(* IEC 61131-3 sources: daoli-st-library/DL_Base (part 18) *)

(* ---- FB_DL_SweepFreqGen.st ---- *)
(*
  Name        : FB_DL_SweepFreqGen
  Category    : DL_Base
  Version     : 1.0.0
  Purpose     : 频率扫描激励发生：线性/对数两模式按起止频率 + 驻留时间表逐段推进，相位逐拍积分输出瞬时频率与相位；/ Frequency sweep excitation generator: linear or logarithmic mode stepping through a dwell-time table between start and stop frequency, with per-scan phase integration
  溯源        : 借 lgf-siggen 的频率发生族待挖组织，clean-room 实现
  Boundary    : ① 起/止频率正域且相等不立（相等退化点频拒绝），越域锁存故障；
                ② 对数扫频禁对零取对数：起频下限 > 0 由正域闸保证（EXP/LN 仅作用于正比值）；
                ③ 相位积分逐拍累加防跳频突跳，相位回卷 2π 用条件减法（禁取模），回卷循环带上限守卫；
                ④ 使能撤除相位保持不归零，bRestart 上升沿显式重启回首段首相位；
                ⑤ 驻留表下标越界钳位（下标域闸）+ 非正驻留钳最小驻留常量；非有限派生频率该拍冻结保持输出；
                ⑥ 本件只出频率/相位激励量，不直接驱动脉冲输出口（属主边界，与 PulseGenerator 职责分立）。
*)
TYPE E_DL_SwpMode :
(
    eLin := 0,                               (* 线性扫频 / Linear sweep *)
    eLog := 10                               (* 对数扫频 / Logarithmic sweep *)
);
END_TYPE

TYPE E_DL_SwpState :
(
    eIdle  := 0,                             (* 未使能（相位保持） / Disabled, phase held *)
    eRun   := 10,                            (* 扫频运行 / Sweeping *)
    eFault := 90                             (* 故障锁存相 / Fault latched *)
);
END_TYPE

TYPE E_DL_SwpCause :
(
    eNone      := 0,                         (* 无故障成因 / No cause *)
    eCfgIllegal:= 1,                        (* 组态非法：频率域/步数/周期越域 / Illegal config *)
    ePhaseBad  := 2                         (* 非法相位兜底 / Illegal phase fallback *)
);
END_TYPE

FUNCTION_BLOCK FB_DL_SweepFreqGen
VAR_INPUT
    fStart  : REAL := 1.0;                   (* 起始频率，域 > 0 且不等于止频 [Hz] / Start frequency *)
    fEnd    : REAL := 100.0;                 (* 结束频率，域 > 0 且不等于起频 [Hz] / Stop frequency *)
    eMode   : E_DL_SwpMode := E_DL_SwpMode.eLin;   (* 扫频模式 / Sweep mode *)
    nSteps  : INT := 8;                      (* 驻留段数，域 2..32 [段] / Dwell step count *)
    aDwell  : ARRAY[1..32] OF TIME;          (* 各段驻留时间表（越界/非正钳位）[ms] / Dwell time table *)
    tScan   : TIME := T#10MS;                (* 扫描周期，域 > T#0S [ms] / Scan period *)
    bRepeat : BOOL := TRUE;                  (* 扫完循环重扫 [-] / Repeat sweep *)
    bEnable : BOOL := TRUE;                  (* 使能（撤除相位保持）[-] / Enable *)
    bRestart: BOOL := FALSE;                 (* 重启命令，上升沿回首段 [-] / Restart command *)
    bReset  : BOOL := FALSE;                 (* 复位命令，上升沿清故障与相位 [-] / Reset command *)
END_VAR
VAR_OUTPUT
    fFreq   : REAL;                          (* 当前瞬时频率出口 [Hz] / Instantaneous frequency outlet *)
    fPhase  : REAL;                          (* 相位累计出口（撤使能保持）[rad] / Phase accumulator outlet *)
    bSweepDone: BOOL;                        (* 单遍扫完脉冲（单拍）[-] / Sweep done pulse *)
    nSegIdx : INT;                           (* 当前段序号 [段] / Current segment index *)
    eState  : E_DL_SwpState;                 (* 状态出口 / State outlet *)
    eCause  : E_DL_SwpCause;                 (* 故障成因出口（R190 归因唯一） / Fault cause outlet *)
    bError  : BOOL;                          (* 故障锁存标志 [-] / Fault latch flag *)
END_VAR
VAR
    _eState : E_DL_SwpState := E_DL_SwpState.eIdle;  (* 内部相位（CASE 唯一写入目标） / Internal phase *)
    _eCause : E_DL_SwpCause := E_DL_SwpCause.eNone;  (* 故障成因锁存量 / Latched cause *)
    rtRestart: R_TRIG;                       (* 重启沿实例，段 0 无条件调用 / Restart edge instance *)
    rtReset : R_TRIG;                        (* 复位沿实例，段 0 无条件调用 / Reset edge instance *)
    _bFault : BOOL;                          (* 故障锁存位 / Latched fault bit *)
    _bCfgBad: BOOL;                          (* 组态非法当拍量 / Illegal config this scan *)
    _bDoneI : BOOL;                          (* 扫完脉冲内部量（统一出口映射，R187） / Done pulse internal *)
    _bFinI  : BOOL;                          (* 派生频率有限性当拍量（边界⑤） / Derived frequency finiteness *)
    _nStepsE: INT;                           (* 钳位后生效段数 [段] / Effective step count *)
    _nSegI  : INT;                           (* 内部当前段序号 [段] / Internal segment index *)
    _fDtSec : REAL;                          (* 扫描周期秒值，域 > eps [s] / Scan period seconds *)
    _fDwellS: REAL;                          (* 当前段驻留秒值（钳位后）[s] / Current dwell seconds *)
    _fTacc  : REAL;                          (* 段内驻留计时累加量 [s] / Dwell time accumulator *)
    _fFreqI : REAL;                          (* 内部瞬时频率中间量 [Hz] / Internal frequency *)
    _fPhaseI: REAL;                          (* 内部相位累计量 [rad] / Internal phase *)
    _fRatio : REAL;                          (* 对数模式频比中间量（恒正）[-] / Log mode ratio *)
    _fWrap  : INT;                           (* 相位回卷守卫计数（防死循环）[次] / Phase wrap guard *)
    _i      : INT;                           (* 驻留表下标中间量 [段] / Dwell table index *)
END_VAR
VAR CONSTANT
    DL_SWP_NMIN  : INT   := 2;               (* 段数下限（边界①域闸配套）[段] / Step count lower bound *)
    DL_SWP_NMAX  : INT   := 32;              (* 段数上限 [段] / Step count upper bound *)
    DL_SWP_EPS   : REAL  := 1.0E-6;          (* 判零容差 [-] / Epsilon *)
    DL_SWP_2PI   : REAL  := 6.2831853;       (* 相位回卷阈（2π 常量）[rad] / Phase wrap threshold *)
    DL_SWP_WRAPMAX: INT  := 64;              (* 相位回卷循环守卫上限（防死循环，边界③）[次] / Wrap loop guard *)
    DL_SWP_TDWMIN: REAL  := 0.01;            (* 最小驻留秒值（非正驻留钳位，边界⑤）[s] / Min dwell seconds *)
END_VAR

(* —— 段 0：当拍判据派生 + 实例无条件刷新（R228A） —— *)
_fDtSec := TIME_TO_LREAL(tScan) / 1000.0;                (* 扫描周期秒化（除子常量 1000） / Scan period seconds *)
_bCfgBad := (fStart <= DL_SWP_EPS) OR (fEnd <= DL_SWP_EPS)              (* 起止频率正域闸（边界①②） / Frequency positive gates *)
            OR (ABS(fStart - fEnd) < DL_SWP_EPS)                        (* 起止相等拒绝（退化点频不立，边界①） / Equal rejected *)
            OR (nSteps < DL_SWP_NMIN) OR (nSteps > DL_SWP_NMAX)         (* 段数域闸 / Step count gate *)
            OR NOT (tScan > T#0S);                                      (* 扫描周期正域闸 / Scan period gate *)
rtRestart(CLK := bRestart);                              (* 重启沿每拍必调 / Restart edge every scan *)
rtReset(CLK := bReset);                                  (* 复位沿每拍必调 / Reset edge every scan *)
_nStepsE := nSteps;                                      (* 生效段数初值 / Effective steps init *)
IF _nStepsE < DL_SWP_NMIN THEN
    _nStepsE := DL_SWP_NMIN;                             (* 段数下限钳位 / Steps lower clamp *)
END_IF
IF _nStepsE > DL_SWP_NMAX THEN
    _nStepsE := DL_SWP_NMAX;                             (* 段数上限钳位 / Steps upper clamp *)
END_IF

(* —— 段 1：单拍量预清零（R107） —— *)
_bDoneI := FALSE;                                        (* 扫完脉冲内部量预清 / Done preset *)
bSweepDone := FALSE;                                     (* 扫完脉冲出口预清 / Done outlet preset *)
_fFreqI := fFreq;                                        (* 频率中间量保持上拍（非有限拍冻结语义，边界⑤） / Frequency hold default *)

(* —— 段 2：复位沿处理（作用域：清故障 + 清相位与段序 + 迁 eIdle，R283 逐项声明） —— *)
IF rtReset.Q THEN
    _bFault := FALSE;                                    (* 清故障锁存 / Clear fault *)
    _eCause := E_DL_SwpCause.eNone;                      (* 清成因 / Clear cause *)
    _fPhaseI := 0.0;                                     (* 清相位累计 / Clear phase *)
    _nSegI := 1;                                         (* 段序回首段 / Segment to first *)
    _fTacc := 0.0;                                       (* 清驻留计时 / Clear dwell timer *)
    fFreq := 0.0;                                        (* 清频率出口 / Clear frequency outlet *)
    fPhase := 0.0;                                       (* 清相位出口 / Clear phase outlet *)
    _eState := E_DL_SwpState.eIdle;                      (* 迁未使能相 / Back to idle *)
END_IF

(* —— 段 3：组态故障锁存（锁存至复位沿，R189） —— *)
IF _bCfgBad AND NOT _bFault THEN
    _bFault := TRUE;                                     (* 锁存故障位 / Latch fault *)
    _eCause := E_DL_SwpCause.eCfgIllegal;                (* 成因：组态非法 / Cause illegal config *)
    _eState := E_DL_SwpState.eFault;                     (* 同步迁故障相 / Migrate to fault *)
END_IF

(* —— 段 4：CASE 主状态机（ELSE 兜底迁 eFault，红线 6） —— *)
CASE _eState OF
    E_DL_SwpState.eIdle:                                 (* 未使能：相位保持不归零（边界④），频率出口确定 0 / Idle *)
        fFreq := 0.0;                                    (* 失能频率出口确定值 / Disabled frequency zero *)
        IF bEnable AND NOT _bFault THEN
            _nSegI := 1;                                 (* 迁入拍段序回首段 / Segment to first *)
            _fTacc := 0.0;                               (* 驻留计时归零 / Dwell timer zero *)
            _eState := E_DL_SwpState.eRun;               (* 进入扫频相 / Enter sweeping *)
        END_IF
    E_DL_SwpState.eRun:                                  (* 扫频相：段推进 + 相位积分 / Sweeping *)
        IF NOT bEnable THEN
            _eState := E_DL_SwpState.eIdle;              (* 失能回未使能（相位保持） / Back to idle *)
        ELSE
            IF rtRestart.Q THEN
                _nSegI := 1;                             (* 显式重启回首段（边界④） / Explicit restart *)
                _fTacc := 0.0;                           (* 驻留计时归零 / Dwell timer zero *)
                _fPhaseI := 0.0;                         (* 重启相位归零 / Phase zero *)
            END_IF
            _i := _nSegI;                                (* 驻留表下标中间量 / Dwell index *)
            IF _i < 1 THEN
                _i := 1;                                 (* 下标下钳（防越界读，边界⑤） / Index lower clamp *)
            END_IF
            IF _i > DL_SWP_NMAX THEN
                _i := DL_SWP_NMAX;                       (* 下标上钳（防越界读，边界⑤） / Index upper clamp *)
            END_IF
            _fDwellS := TIME_TO_LREAL(aDwell[_i]) / 1000.0;   (* 驻留秒化（除子常量 1000） / Dwell seconds *)
            IF _fDwellS < DL_SWP_TDWMIN THEN
                _fDwellS := DL_SWP_TDWMIN;               (* 非正/过小驻留钳最小值（边界⑤） / Dwell clamp *)
            END_IF
            IF _fDtSec > DL_SWP_EPS THEN                 (* 周期秒值有效才推进（防除零/防零步进） / Period gate *)
                IF eMode = E_DL_SwpMode.eLog THEN
                    _fRatio := fEnd / fStart;            (* 对数频比（分子分母均过正域闸，边界②） / Log ratio *)
                    _fFreqI := fStart * EXP(LN(_fRatio) * INT_TO_REAL(_nSegI - 1) / INT_TO_REAL(_nStepsE - 1));   (* 几何步进频率（除子 = 段数-1 >= 1） / Geometric frequency *)
                ELSE
                    _fFreqI := fStart + (fEnd - fStart) * INT_TO_REAL(_nSegI - 1) / INT_TO_REAL(_nStepsE - 1);    (* 线性步进频率（除子 >= 1） / Linear frequency *)
                END_IF
                _bFinI := (_fFreqI = _fFreqI) AND ((_fFreqI - _fFreqI) = (_fFreqI - _fFreqI));   (* 派生频率有限性闸（边界⑤） / Derived finiteness gate *)
                IF _bFinI THEN
                    _fPhaseI := _fPhaseI + DL_SWP_2PI * _fFreqI * _fDtSec;   (* 相位逐拍积分防跳频突跳（边界③） / Phase integrate *)
                    _fWrap := 0;                         (* 回卷守卫计数清零 / Wrap guard clear *)
                    WHILE (_fPhaseI >= DL_SWP_2PI) AND (_fWrap < DL_SWP_WRAPMAX) DO   (* 条件减法回卷（禁取模，边界③） / Conditional wrap *)
                        _fPhaseI := _fPhaseI - DL_SWP_2PI;   (* 相位减 2π / Phase minus 2 pi *)
                        _fWrap := _fWrap + 1;            (* 守卫计数递进 / Guard advance *)
                    END_WHILE
                    fFreq := _fFreqI;                    (* 频率出口（有限拍派生） / Frequency outlet *)
                    fPhase := _fPhaseI;                  (* 相位出口 / Phase outlet *)
                    _fTacc := _fTacc + _fDtSec;          (* 段内驻留计时累加 / Dwell timer advance *)
                    IF _fTacc >= _fDwellS THEN           (* 驻留满迁下一段 / Dwell elapsed *)
                        _fTacc := 0.0;                   (* 驻留计时重置（R227） / Dwell timer reset *)
                        _nSegI := _nSegI + 1;            (* 段序净额 +1 / Segment advance *)
                        IF _nSegI > _nStepsE THEN        (* 末段完成 / Last segment done *)
                            _bDoneI := TRUE;             (* 扫完脉冲内部置位（R187） / Done internal *)
                            IF bRepeat THEN
                                _nSegI := 1;             (* 循环重扫回首段 / Repeat to first *)
                            ELSE
                                _nSegI := _nStepsE;      (* 单遍模式停末段（频率保持） / Hold last segment *)
                            END_IF
                        END_IF
                    END_IF
                END_IF                                   (* 非有限拍：频率/相位冻结保持上拍（边界⑤） *)
            END_IF
            nSegIdx := _nSegI;                           (* 当前段序号出口 / Segment index outlet *)
        END_IF
    E_DL_SwpState.eFault:                                (* 故障相：冻结保持末值，仅复位沿出 / Fault *)
        ;                                                (* 锁存回放（R28） / Replay from latch *)
    ELSE                                                 (* 非法相位兜底迁安全态 / Illegal phase fallback *)
        _eState := E_DL_SwpState.eFault; _bFault := TRUE;    (* 迁故障相 + 同步锁存 / To fault and latch *)
        _eCause := E_DL_SwpCause.ePhaseBad;              (* 成因：非法相位 / Cause illegal phase *)
END_CASE

(* —— 段 5：出口映射（内部 _b* → 输出单拍，R187；名实双出口，R191） —— *)
bSweepDone := _bDoneI;                                   (* 扫完脉冲单拍出口 / Done pulse outlet *)
bError := _bFault;                                       (* 故障标志镜像 / Fault flag mirror *)
eState := _eState;                                       (* 状态出口 / State outlet *)
eCause := _eCause;                                       (* 成因出口 / Cause outlet *)
END_FUNCTION_BLOCK

(* ---- FB_DL_TimerFailSafe.st ---- *)
(*
  ==================================================================
  组件名 Component  : FB_DL_TimerFailSafe
  分类   Category   : DL_Base
  复杂度 Complexity  : 轻
  版本   Version    : 1.0.0
  功能   Purpose    : 安全侧定时器。接通延时输出 bOut；当输出持续时长超过
                      tMaxHold 看门狗窗时自动回安全态 FALSE 并锁存 bTimedOut，
                      解除路径 = bIn 断电或 bReset 上升沿。安全侧赋值单点完成
                      （bOut := tonDelay.Q AND NOT _bLatch），不受本闸判定量
                      污染；与 FB_DL_ExtendedTimer 通用四模式分工互引。
  来源   Source     : T0-iec-std-wrapper（T0-2 定时器安全语义扩展）
  溯源   Origin     : IEC 61131-3 TON 标准语义的安全包装，clean-room 自研实现，
                      未复制任何厂商私有库源码。
  平台   Platform   : 纯 IEC 61131-3（Standard.library: TON / R_TRIG，无私有库）
  分工声明 Split     : 与 FB_DL_ExtendedTimer 分工——后者做通用四模式定时，
                      本件只做安全侧超时自动回退封装。
  作者   Author     : 道莅代码库 · PLC 编程专家（R59）
  ------------------------------------------------------------------
  边界 Boundary     :
                      一 安全语义：bOut 唯一赋值点为统一出口，锁存期强制 FALSE
                         （安全态），锁存解除后须 bIn 重新接通才重新计时；
                      二 组态域：tOnDelay / tMaxHold 由调用方保证为正时长，
                         本件不做二次钳制；
                      三 定时器与沿检测全部段 0 无条件周期刷新（R7）；
                      四 无全局变量、无外部变量声明、无物理地址寻址。
  修订记录 Revision  :
    2026-11-21  v1.0.0  R59 首版（批 1 · 序号 1）
  ==================================================================
*)

FUNCTION_BLOCK FB_DL_TimerFailSafe
VAR_INPUT
    bIn       : BOOL := FALSE;  // 定时条件输入，TRUE = 请求延时接通 [-] / the timing condition input, true = the on delay requested
    tOnDelay  : TIME := T#2S;   // 接通延时整定 [毫秒] / the on delay setting [millisecond]
    tMaxHold  : TIME := T#60S;  // 输出最大允许持续时长，超过自动安全态 [毫秒] / the max allowed hold duration, safe state beyond [millisecond]
    bReset    : BOOL := FALSE;  // 超时锁存复位，上升沿生效 [-] / the timeout latch reset, rising edge effective
END_VAR
VAR_OUTPUT
    bOut      : BOOL := FALSE;  // 安全侧定时输出，超时自动回 FALSE [-] / the safety side timed output, safe false on timeout
    bRun      : BOOL := FALSE;  // 延时计时进行指示 [-] / the delay timing in progress indicator
    bTimedOut : BOOL := FALSE;  // 超时锁存指示，解除 = bIn 断电或复位沿 [-] / the timeout latch indicator, released by input drop or reset edge
    bError    : BOOL := FALSE;  // 预留故障位（本件无浮点运算，恒常假）[-] / the reserved fault bit, constant false in this block
END_VAR
VAR
    _bInit   : BOOL := FALSE; // 首拍初始化标志（R310，真实使用：首拍强制安全态预置）/ the first scan flag, real use, the safe preset on first scan
    _bLatch  : BOOL := FALSE; // 超时锁存位（安全态保持源，区分于实时镜像 bTimedOut）/ the timeout latch bit, the safe state source
    rtReset  : R_TRIG;        // 复位沿检测，段 0 无条件刷新 / the reset edge, refreshed unconditionally at segment 0
    tonDelay : TON;           // 接通延时器，段 0 无条件刷新 / the on delay timer, refreshed unconditionally
    tonHold  : TON;           // 持续时长看门狗，段 0 无条件刷新 / the hold watchdog timer, refreshed unconditionally
END_VAR

// 段 0｜定时器与沿检测无条件周期刷新（禁入分支，R7）/ segment 0, the unconditional refresh
rtReset(CLK := bReset); // 复位沿 / the reset edge
tonDelay(IN := bIn AND (NOT _bLatch), PT := tOnDelay); // 接通延时，锁存期不计时 / the on delay, not timing while latched
tonHold(IN := tonDelay.Q AND (NOT _bLatch), PT := tMaxHold); // 持续看门狗，仅在输出成立期计时 / the hold watchdog, timing only while the output stands

// 段 1｜首拍初始化（R310 真实使用路径）：强制安全态预置 / segment 1, the first scan init, the safe preset
IF NOT _bInit THEN // 首拍一拍 / the first scan
    _bInit := TRUE; // 置首拍标志 / raise the first scan flag
    _bLatch := FALSE; // 锁存清零（编译缺省之上的显式安全预置）/ clear the latch explicitly
    bOut := FALSE; // 输出强制安全态 / force the output safe
END_IF

// 段 2｜超时锁存与解除（锁存解除路径 = bIn 断电沿或 bReset 上升沿，双路径可达，R188）/ segment 2, the timeout latch and release
IF tonHold.Q THEN // 看门狗窗到期：超时锁存 / the watchdog expired, latch the timeout
    _bLatch := TRUE; // 置超时锁存 / raise the timeout latch
END_IF
IF (NOT bIn) OR rtReset.Q THEN // 条件断电或复位沿 / the condition dropped or the reset edge
    _bLatch := FALSE; // 解除锁存（解除后再接通需重新计时）/ release the latch
END_IF

// 段 3｜统一出口：安全侧赋值单点完成（判定量 bIn 只经 tonDelay.Q 进入，不被闸判定量污染，边界一）/ segment 3, the unified outlet
bOut := tonDelay.Q AND (NOT _bLatch); // 输出 = 延时到 且 未超时锁存 / the output, delayed and not latched
bRun := tonDelay.IN; // 计时进行镜像 / the timing in progress mirror
bTimedOut := _bLatch; // 超时指示与锁存位同源（R191 名实双出口）/ the timeout indicator shares the latch
END_FUNCTION_BLOCK

(* ---- FB_DL_TimeWindowCheck.st ---- *)
(*==============================================================================
 * 组件名称 (Component)  : FB_DL_TimeWindowCheck
 * 所属子库 (Sublibrary) : DL_Base
 * 当前版本 (Version)    : 1.0.0
 * 兼容性   (Platform)   : CODESYS 3.5 / TwinCAT 3 / 汇川 InoProShop / Machine Expert
 *                         仅依赖 Standard.library（R_TRIG / MIN），零厂商方言
 * 分类     (Category)   : 功能块（FUNCTION_BLOCK）· 每日时间窗判定 · Level 0 DL_Base 补强件
 * 功能描述 (Function)   : 每日时间窗单一语义判定块（LGF mode 巨无霸反例的落实：
 *                         不设 MODE 参数，每周/每月/每年窗按矩阵扩产规则拆独立
 *                         块）。判定 = 本日总使能 AND 星期表当日位 AND 时刻窗。
 *                         时刻窗支持跨零点（如 22:00→06:00：t≥开 OR t<关）；
 *                         开=关视为 24h 全开（语义见段内注释）。窗口开/闭沿
 *                         单发脉冲供启停设备一次触发。当前时刻/星期由引脚注入
 *                         （零全局耦合红线：禁读 CPU 本地钟），典型与
 *                         FC_DL_DayOfWeekCalc 输出直连。
 * 开源溯源 (Origin)     : 来源标签 lgf-datetime（Siemens LGF V5.2.1 · 3.1 Date
 *                         and timer operations 章 定时开关族）。仅借鉴每日窗/
 *                         跨零点判定与星期使能表的公开行为语义；去 mode 巨无霸
 *                         化（单一语义拆块）、去 CPU 钟耦合（时间引脚注入）均
 *                         为本库独立设计决策，clean-room 重写，未复制任何源码行。
 * 本文件内含       : FUNCTION_BLOCK FB_DL_TimeWindowCheck
 * 依赖     (Depends)    : Standard.library: R_TRIG / MIN；建议上游搭配
 *                          FC_DL_DayOfWeekCalc（ISO 序星期源，引脚注入）。
 *                          不引用 DL_ 内其他实现文件。
 * 故障码表 (Error codes) : 16#0001_0202【信息级】时刻/星期参数越界（当前时刻越
 *                          界按 FALSE 处理；窗口参数越界按钳位后照常计算），
 *                          不置任何故障位（本块无故障锁存位）；0 = 无。沿用
 *                          DL_Base 既有 16#0001_xxxx 段，与 VERSION.md 故障码
 *                          表无冲突。
 * 【规格偏离留档 / R11 Deviation register】
 *   D1 规格 §4.2 引脚表未提供星期索引注入引脚，aWeekdayEnable[1..7] 表在块内
 *      无法自索引（时刻引脚不含日期信息）；按 R11 留档新增输入引脚
 *      uWeekdayNow : USINT := 1（当前星期注入，ISO 序 1=周一..7=周日，与
 *      §4.1 FC_DL_DayOfWeekCalc 输出同序同域），越界不读表并置信息级码。
 *   D2 规格引脚表 bReset 注释为「—」：本块定义其语义为上升沿清除当拍信息级码
 *      并强制重新评估窗口（日切换后防陈旧码残留），不影响窗口判定结果本身。
 * 红线自检 (Redline)    : R1 ✓ 零全局变量表与外部变量引用 ｜ R2 ✓ 零物理 IO 地址直写
 *                         R3 ✓ 纯 IEC 61131-3 ｜ R4 ✓ 越界防御+分钟折算 UINT 扩宽防溢出
 *                         R5 ✓ 全变量中英双语同行注释 ｜ R6 不适用（组合逻辑+沿检测，无状态机）
 *                         R7 ✓ 三个 R_TRIG 实例主体无条件周期刷新（严禁入分支）
 * 修订历史 (Revision)   :
 *   2026-11-15  v1.0.0  首版入库 · Round 05 · 泳道 B · 契约出处 ROUND_PLAN_R5 §4.2
 * 验收向量 (Acceptance) :
 *   V1 同日窗：On=08:00 / Off=18:00，Now=12:00 → bInWindow=TRUE；Now=07:59 /
 *      18:00 → FALSE（左闭右开）
 *   V2 跨零点窗：On=22:00 / Off=06:00，Now=23:30 或 05:59 → TRUE；Now=06:00 →
 *      FALSE；Now=21:59 → FALSE
 *   V3 24h 窗：On=Off=08:00 → 任意时刻 bInWindow=TRUE（开=关全开语义）
 *   V4 星期表：uWeekdayNow=6（周六）且 aWeekdayEnable[6]=FALSE → 不在窗，其余
 *      条件不影响；uWeekdayNow=0 或 8 → 信息级 0001_0202 且按不在窗处理
 *   V5 时刻越界：uHourNow=24 → bInWindow=FALSE + 0001_0202（当前时刻越界按
 *      FALSE 处理）；uHourOn=25 → 钳位 23 后照常计算 + 0001_0202（信息级钳位）
 *   V6 沿单发：V1 场景下 Now 由 07:59 → 08:00 当拍 bPulseOnWindowOpen=TRUE 单发；
 *      18:00 当拍 bPulseOnWindowClose=TRUE 单发
 *   V7 复位沿：越界码出现后 bReset 上升沿当拍 uErrorId 清零（触发实例无条件刷新）
 *============================================================================*)

(*==============================================================================
 * 功能块: FB_DL_TimeWindowCheck
 * 调用约定: 每个扫描周期无条件调用一次；三个 R_TRIG 实例在主体无条件周期刷新，
 *           严禁移入 IF/CASE 分支（R7）。时刻/星期由调用方每拍注入。
 *============================================================================*)
FUNCTION_BLOCK FB_DL_TimeWindowCheck
VAR_INPUT
    uHourNow        : USINT;                // 当前时刻-时（Injected local time hour）[h] 0..23，越界按不在窗处理（禁读 CPU 钟，公约 0.9）
    uMinNow         : USINT;                // 当前时刻-分（Injected local time minute）[min] 0..59
    bEnableDay      : BOOL := TRUE;         // 本日窗总使能（Day window enable），FALSE 时恒不在窗
    aWeekdayEnable  : ARRAY[1..7] OF BOOL;  // 周一~周日各日使能表（Weekday enable table），索引 1=周一（ISO 序，与 FC_DL_DayOfWeekCalc 一致）
    uWeekdayNow     : USINT := 1;           // 【偏离 D1 新增】当前星期注入（Injected weekday）1=周一..7=周日（ISO 序），越界不读表
    uHourOn         : USINT := 6;           // 窗口开启-时（Window on hour）[h] 0..23，越界钳位后照算（公约 0.2）
    uMinOn          : USINT := 0;           // 窗口开启-分（Window on minute）[min] 0..59
    uHourOff        : USINT := 22;          // 窗口关闭-时（Window off hour）[h] 0..23，支持跨零点（如 22:00→06:00）
    uMinOff         : USINT := 0;           // 窗口关闭-分（Window off minute）[min] 0..59
    bReset          : BOOL := FALSE;        // 复位（Reset）上升沿：清除当拍信息级码并重新评估（偏离 D2）
END_VAR
VAR_OUTPUT
    bInWindow           : BOOL;             // 当前处于窗口内（In window）= 本日使能 AND 星期位 AND 时刻窗
    bPulseOnWindowOpen  : BOOL;             // 窗口开启沿单发（Window open edge），TRUE 持续一拍
    bPulseOnWindowClose : BOOL;             // 窗口关闭沿单发（Window close edge），TRUE 持续一拍
    uErrorId            : UDINT;            // 信息级码（Info code）16#0001_0202 = 时刻/星期越界；0 = 无
END_VAR
VAR
    fbTrigReset     : R_TRIG;               // 复位信号上升沿检测实例（Reset edge detector）
    fbTrigOpen      : R_TRIG;               // 窗口开启沿检测实例（Window open edge detector），CLK = bInWindow
    fbTrigClose     : R_TRIG;               // 窗口关闭沿检测实例（Window close edge detector），CLK = NOT bInWindow
    uHourOnC        : USINT;                // 钳位后开启-时（Clamped on hour）[h] 0..23
    uMinOnC         : USINT;                // 钳位后开启-分（Clamped on minute）[min] 0..59
    uHourOffC       : USINT;                // 钳位后关闭-时（Clamped off hour）[h] 0..23
    uMinOffC        : USINT;                // 钳位后关闭-分（Clamped off minute）[min] 0..59
    uNowMin         : UINT;                 // 当前时刻折算分钟（Now in minutes）0..1439，USINT 域乘法越界防御
    uOnMin          : UINT;                 // 开窗时刻折算分钟（On time in minutes）0..1439
    uOffMin         : UINT;                 // 关窗时刻折算分钟（Off time in minutes）0..1439
    bTimeNowOk      : BOOL;                 // 当前时刻有效性（Now time valid）
    bWinParamOk     : BOOL;                 // 窗口参数有效性（Window params valid）
    bWeekdayOk      : BOOL;                 // 星期索引有效性（Weekday index valid）
    bTimeInWin      : BOOL;                 // 时刻窗判定结果（Time-in-window result）
    bDayOk          : BOOL;                 // 日使能合成结果（Day-enable result）
END_VAR

// -----------------------------------------------------------------------------
// 段 1｜边沿实例无条件周期刷新（R7 红线：严禁移入 IF/CASE 分支）
// -----------------------------------------------------------------------------
fbTrigReset(CLK := bReset);                 // 复位沿检测

// -----------------------------------------------------------------------------
// 段 2｜有效性判定与信息级码准备（信息级 0001_0202 只进 uErrorId，本块无故障位）
// -----------------------------------------------------------------------------
uErrorId := 16#0000_0000;                   // 每拍重算信息级码
bTimeNowOk  := (uHourNow <= 23) AND (uMinNow <= 59);               // 当前时刻域检查
bWinParamOk := (uHourOn <= 23) AND (uMinOn <= 59)
            AND (uHourOff <= 23) AND (uMinOff <= 59);          // 窗口参数域检查
bWeekdayOk  := (uWeekdayNow >= 1) AND (uWeekdayNow <= 7);      // 星期索引域检查（ISO 1..7）
IF NOT bTimeNowOk THEN
    uErrorId := 16#0001_0202;               // 当前时刻越界：按不在窗处理（引脚注释基线）
END_IF
IF NOT bWinParamOk THEN
    uErrorId := 16#0001_0202;               // 窗口参数越界：钳位后照常计算（公约 0.2）
END_IF
IF NOT bWeekdayOk THEN
    uErrorId := 16#0001_0202;               // 星期索引越界：不读表，按不在窗处理
END_IF

// -----------------------------------------------------------------------------
// 段 3｜窗口参数钳位（信息级钳位，钳位后继续计算，不中断扫描）
// -----------------------------------------------------------------------------
uHourOnC  := MIN(uHourOn, 23);              // 开启-时钳位 [h]
uMinOnC   := MIN(uMinOn, 59);               // 开启-分钳位 [min]
uHourOffC := MIN(uHourOff, 23);             // 关闭-时钳位 [h]
uMinOffC  := MIN(uMinOff, 59);              // 关闭-分钳位 [min]

// -----------------------------------------------------------------------------
// 段 4｜分钟折算（USINT×60 最大 1380 超 USINT 域，先扩宽 UINT 再运算防越界）
// -----------------------------------------------------------------------------
uOnMin := uHourOnC;                         // USINT → UINT 隐式扩宽
uOnMin := (uOnMin * 60) + uMinOnC;          // 开窗分钟 [min] 0..1439
uOffMin := uHourOffC;                       // USINT → UINT 隐式扩宽
uOffMin := (uOffMin * 60) + uMinOffC;       // 关窗分钟 [min] 0..1439
IF bTimeNowOk THEN
    uNowMin := uHourNow;                    // USINT → UINT 隐式扩宽
    uNowMin := (uNowMin * 60) + uMinNow;    // 当前分钟 [min] 0..1439
ELSE
    uNowMin := 0;                           // 时刻越界：折算值弃用，结果由 bTimeNowOk 门控
END_IF

// -----------------------------------------------------------------------------
// 段 5｜时刻窗判定（跨零点支持；开=关视为 24h 全开——语义：本日整日放行）
// -----------------------------------------------------------------------------
IF uOnMin > uOffMin THEN
    bTimeInWin := (uNowMin >= uOnMin) OR (uNowMin < uOffMin);   // 跨零点窗：t≥开 OR t<关（如 22:00→06:00）
ELSIF uOnMin < uOffMin THEN
    bTimeInWin := (uNowMin >= uOnMin) AND (uNowMin < uOffMin);  // 同日窗：开≤t<关（左闭右开）
ELSE
    bTimeInWin := TRUE;                                          // 开=关：24h 全开（每日窗单一语义特例）
END_IF

// -----------------------------------------------------------------------------
// 段 6｜日使能合成（星期越界不读表，防数组越界，R4）
// -----------------------------------------------------------------------------
IF bWeekdayOk THEN
    bDayOk := bEnableDay AND aWeekdayEnable[uWeekdayNow];       // 总使能 AND 当日星期位（索引 1..7 已校验）
ELSE
    bDayOk := FALSE;                        // 星期索引越界：按不在窗处理
END_IF

// -----------------------------------------------------------------------------
// 段 7｜总判定：当前时刻越界按 FALSE 处理；窗口参数已钳位故不再门控结果
// -----------------------------------------------------------------------------
bInWindow := bDayOk AND bTimeNowOk AND bTimeInWin;              // 在窗 = 日使能 AND 时刻有效 AND 时刻窗

// -----------------------------------------------------------------------------
// 段 8｜窗口开/闭沿单发（实例无条件周期刷新，沿输出各持续一拍）
// -----------------------------------------------------------------------------
fbTrigOpen(CLK := bInWindow);               // 开启沿检测
fbTrigClose(CLK := NOT bInWindow);          // 关闭沿检测（取反 CLK）
bPulseOnWindowOpen  := fbTrigOpen.Q;        // 开启沿单发输出
bPulseOnWindowClose := fbTrigClose.Q;       // 关闭沿单发输出

// -----------------------------------------------------------------------------
// 段 9｜复位沿消费：清除当拍信息级码（触发实例已在段 1 无条件刷新，偏离 D2）
// -----------------------------------------------------------------------------
IF fbTrigReset.Q THEN
    uErrorId := 16#0000_0000;               // 复位沿当拍清信息级码（下一拍重新评估）
END_IF

END_FUNCTION_BLOCK

(* ---- FB_DL_TofEx.st ---- *)
(*==============================================================================
 * 组件名称 (Component)  : FB_DL_TofEx
 * 所属子库 (Sublibrary) : DL_Base
 * 当前版本 (Version)    : 1.0.0
 * 兼容性   (Platform)   : CODESYS 3.5 / TwinCAT 3 / 汇川 InoProShop / Machine Expert
 *                         仅依赖 Standard.library（TOF），零厂商方言
 * 功能描述 (Function)   : 断开延时定时器防御包装。内部委托 IEC 61131-3 标准 TOF
 *                         实例完成计时内核，外围提供 PT 负值钳位、首扫语义统一
 *                         （首扫 bIN=FALSE 时 bQ 必为 FALSE）与跨段语义直通。
 * 溯源     (Origin)     : IEC 61131-3 标准语义的道莅防御性实现
 *                         （接口语义由 IEC 61131-3 定义，clean-room 重写，
 *                         参考公开标准条款）
 * 码位     (Diag Codes) : 信息级占用区间 16#0001_0150（本件独占，仅此一码）
 *                         16#0001_0150 = tPT 为负值，已钳位为 T#0s（信息级，
 *                         钳位属正常防御行为，不置故障）
 * 类型裁定 (Type Note)  : 码位段 16#0001_xxxx 为全库共享 32 位段，WORD 容量不足，
 *                         故 uDiag 采用 UDINT 承载（与库内 uErrorId : UDINT 惯例一致）
 * 依赖     (Depends)    : 无 DL_ 内部依赖；Standard.library: TOF
 * 红线自检 (Redline)    : R1 ✓ 零全局变量与外部变量引用 ｜ R2 ✓ 零物理 IO 地址直写
 *                         R3 ✓ 纯 IEC 61131-3 ｜ R4 ✓ PT 钳位+除零/越界无涉
 *                         R5 ✓ 全变量中英双语同行注释 ｜ R6 N/A（无顺序状态机，见下）
 *                         R7 ✓ TOF 实例主体无条件周期刷新
 * 说明     (Note)       : R6 标注 N/A —— 本组件为单步延时逻辑，不存在顺序状态机，
 *                         无 CASE 可写；唯一状态即"延时中/直通"，以本节说明
 *                         替代 ELSE 兜底，符合"无状态机则标注 N/A"口径。
 * 防御行为声明 (Defense): ① tPT < T#0s 时钳位为 T#0s 并置信息码 16#0001_0150
 *                           （部分平台负 TIME 行为未定义，本库统一钳 0）；
 *                         ② 首扫语义统一：首扫 bIN=FALSE 时 bQ 必为 FALSE、tET=T#0s
 *                           ——由内建 TOF 标准行为（Q 随 IN 直通 + 断开延时）保证，
 *                           部分平台首扫假触发差异在包装层被标准实例天然屏蔽；
 *                         ③ bIN 接通当拍 tET 归零、bQ 立即 TRUE（IEC TOF 标准语义，
 *                           包装层不重实现）。
 * 修订历史 (Revision)   :
 *   2026-11-16  v1.0.0  首版入库（R14 批 2 · T0 快车道）
 *============================================================================*)
FUNCTION_BLOCK FB_DL_TofEx
VAR_INPUT
    bIN : BOOL;   // 定时输入，TRUE 直通输出，FALSE 起断开延时 / Timing input, TRUE passes through, FALSE starts the off-delay
    tPT : TIME;   // 预置延时 [ms]，负值将被钳位为 T#0s / Preset delay [ms], negative values are clamped to T#0s
END_VAR
VAR_OUTPUT
    bQ    : BOOL;   // 输出，bIN 断开并持续 tPT 后变 FALSE / Output, goes FALSE after bIN held FALSE for tPT
    tET   : TIME;   // 已计时 [ms]，bIN 接通当拍归零 / Elapsed time [ms], zeroed on the scan bIN rises
    uDiag : UDINT;  // 诊断字，16#0001_0150=tPT 负值已钳 0，0=无诊断事件 / Diag word, 16#0001_0150=negative tPT clamped to 0, 0=no diag event
END_VAR
VAR
    fbTof    : TOF;   // 内建断开延时实例，承担计时内核 / Built-in TOF instance, owns the timing kernel
    tPTClamp : TIME;  // 钳位后的预置延时 [ms]，喂给内建实例 / Clamped preset delay [ms], fed to the built-in instance
    xInit    : BOOL;  // 首扫初始化标志，FALSE=尚未完成上电初始化 / First-scan init flag, FALSE = power-on init not yet done
END_VAR

(*------------------------------------------------------------------------------
 * 段 1｜首扫初始化（历史教训④口径）：置于逻辑最前，首扫不产假 bQ
 *      First-scan init (lesson 4): placed at the very front, no false bQ on first scan
 *-----------------------------------------------------------------------------*)
IF NOT xInit THEN
    xInit    := TRUE;    // 置初始化完成标志 / Mark init as done
    tPTClamp := T#0s;    // 首扫钳位值归零，避免未初始化喂入 / Zero the clamp value on first scan, no uninitialized feed
    uDiag    := 16#0000_0000;  // 首扫诊断字清零 / Clear diag word on first scan
END_IF

(*------------------------------------------------------------------------------
 * 段 2｜PT 域校验与钳位：负 TIME 在部分平台行为未定义，统一钳 0 并置信息码；
 *      写入点排序审计（历史教训⑦）：本件诊断字仅有"置码/清码"单一分支对，
 *      无复位类与置位类竞态，排序安全
 *      PT domain check and clamp: negative TIME is undefined on some platforms,
 *      unified clamp to 0 with an informational code
 *-----------------------------------------------------------------------------*)
IF tPT < T#0s THEN
    tPTClamp := T#0s;        // 负值钳位为 0 [ms] / Clamp negative to 0 [ms]
    uDiag    := 16#0001_0150;  // 信息码：PT 负值已钳 0 / Informational: negative PT clamped to 0
ELSE
    tPTClamp := tPT;         // 域内直通 / In-domain pass-through
    uDiag    := 16#0000_0000;  // 无诊断事件，清码 / No diag event, clear code
END_IF

(*------------------------------------------------------------------------------
 * 段 3｜无条件刷新区（红线 R7）：TOF 实例严禁进入任何 IF / CASE 分支；
 *      首扫 bIN=FALSE → bQ=FALSE 与"接通当拍 ET 归零"均由内建标准语义保证
 *      Unconditional refresh zone (red line R7): no instance call inside IF / CASE;
 *      first-scan bQ=FALSE with bIN=FALSE and ET zeroing on bIN rise are both
 *      guaranteed by the built-in TOF standard behavior
 *-----------------------------------------------------------------------------*)
fbTof(IN := bIN, PT := tPTClamp);  // 每扫描周期无条件喂入输入与钳位后 PT / Feed input and clamped PT unconditionally every scan

(*------------------------------------------------------------------------------
 * 段 4｜输出直通：bQ/tET 逐拍镜像内建实例输出，包装层不重实现计时内核
 *      Output pass-through: bQ/tET mirror the built-in outputs scan by scan;
 *      the wrapper never re-implements the timing kernel
 *-----------------------------------------------------------------------------*)
bQ  := fbTof.Q;   // 输出直通 / Output pass-through
tET := fbTof.ET;  // 已计时 [ms] 直通 / Elapsed time [ms] pass-through
END_FUNCTION_BLOCK

(* ---- FB_DL_ToggleButtonBank.st ---- *)
(*
  FB_DL_ToggleButtonBank  —  多路启停按钮组解算 / Multi-channel toggle button bank solver
  分类 Category : DL_Base
  码位 Code     : 16#01_0_01
  版本 Version  : 1.0.0
  来源 Source   : t1-5-tcopen — IEC 61131-3 标准语义的道莅防御性实现
  溯源 Origin   : TCopen 按钮组/选择器公开语义借鉴，clean-room 实现，未复制任何源码行
  功能 Function : 1) 三种解算模式：Toggle 单按钮逐通道翻转锁存 / SingleAct 双按钮点动直通 / Selector3 三位置选择互斥；
                  2) Selector3 通道互斥：新通道置位时旧通道清零；同拍多键按「低通道号优先」并置信息码（不静默双通）；
                  3) 失电来电恢复策略 eRestorePolicy：Hold 保持（RETAIN 语义由上层承载）/ Reset 全清 / Pulse 上电首拍单周期 TRUE；
                  4) nActiveChannel 输出当前活动通道（0 = 无，1..n = 最低活动通道号，Selector3 即唯一互斥通道）。
  边界 Boundary : ① uChannelCount = 0 或 > nMaxCh 判组态错 bCfgFault，全输出 FALSE（安全侧）；
                  ② 8 路 R_TRIG 在主周期无条件刷新（调用语句不置于 IF/CASE 内，R182）；
                  ③ SingleAct 点动直通不锁存：输出 = 按钮实时电平（松开即断，无保持）；
                  ④ 解除式自证：bCfgFault 解除 = 下一拍 uChannelCount 落回合法域（每拍重算，无锁存）；
                  ⑤ Pulse 脉冲语义：仅上电首拍 abOut 全 TRUE 一个 PLC 周期，第二拍起恢复正常解算（注释标明，防误用为持续使能）。
  依赖 Depends  : 仅 Standard.library（R_TRIG）；枚举 E_DL_BtnMode / E_DL_RestorePolicy 随本件发布
  码表 Error codes（本件格 01_0_01，子码步进 +0x100）:
    16#0001_0101 信息级：Selector3 同拍多键，低通道号优先（不置故障）
    16#0001_0201 故障级：组态非法 uChannelCount = 0 或超数组上界
    16#0001_0301 信息级：Pulse 恢复策略上电首拍单周期脉冲（不置故障）

  修订历史 Revision :
    2026-11-18  v1.0.0  R38 首版
*)

TYPE E_DL_BtnMode :
(
    eToggle    := 0,   // 单按钮翻转锁存 / Single-button toggle with latch
    eSingleAct := 1,   // 点动直通（不锁存）/ Momentary passthrough, no latch
    eSelector3 := 2    // 三位置选择互斥 / Three-position selector, mutually exclusive
);
END_TYPE

TYPE E_DL_RestorePolicy :
(
    eHold  := 0,   // 上电保持断电前状态（RETAIN 由上层承载）/ Hold pre-power-loss state, retainment owned upstream
    eReset := 1,   // 上电全清零 / Clear all outputs at power-up
    ePulse := 2    // 上电首拍单周期 TRUE / Single-scan TRUE pulse at power-up
);
END_TYPE

FUNCTION_BLOCK FB_DL_ToggleButtonBank
VAR_INPUT
    abBtn          : ARRAY[0..7] OF BOOL;   // 按钮输入组 [0..nMaxCh-1] / Button inputs
    uChannelCount  : INT;                   // 有效通道数 [路]，域 1..nMaxCh / Valid channel count
    eMode          : E_DL_BtnMode;          // 解算模式 / Solver mode
    eRestorePolicy : E_DL_RestorePolicy;    // 失电来电恢复策略 / Power-restore policy
END_VAR
VAR_OUTPUT
    abOut          : ARRAY[0..7] OF BOOL;   // 通道输出组 / Channel outputs
    nActiveChannel : INT;                   // 活动通道号（0 = 无，1..n 最低活动）/ Active channel, 0 = none
    bCfgFault      : BOOL;                  // 组态非法（每拍重算）/ Configuration fault, recomputed
    nErrId         : UDINT;                 // 事件码，0 = 无事件 / Event code, 0 = none
END_VAR
VAR
    artBtn     : ARRAY[0..7] OF R_TRIG;     // 逐通道按钮上升沿，段 0 无条件刷新 / Per-channel rising edges
    _abState   : ARRAY[0..7] OF BOOL;       // Toggle 模式锁存状态 / Toggle latched states
    _bFirstScan: BOOL := TRUE;              // 上电首拍标志 / First-scan-after-power-up flag
    _bSimulKey : BOOL;                      // 同拍多键标志（本拍重算）/ Simultaneous keys flag
    _k         : INT;                       // 循环计数器 / Loop counter
END_VAR
VAR CONSTANT
    nMaxCh : INT := 8;                      // 数组上界 [路] / Array upper bound
END_VAR

(* —— 段 0：R_TRIG 无条件周期刷新（R182：调用语句不得置于 IF/CASE 内） —— *)
FOR _k := 0 TO (nMaxCh - 1) DO
    artBtn[_k](CLK := abBtn[_k]);           // 逐通道上升沿，每拍必调
END_FOR

(* —— 段 1：单拍量预清零 —— *)
nErrId     := 16#0000_0000;               // 事件码缺省无事件
_bSimulKey := FALSE;                      // 多键标志预清零
FOR _k := 0 TO (nMaxCh - 1) DO
    abOut[_k] := FALSE;                   // 输出缺省 FALSE（安全侧缺省，段 4 单点置位）
END_FOR
nActiveChannel := 0;                      // 活动通道缺省无

(* —— 段 2：组态域闸（uChannelCount 全覆盖，每拍重算） —— *)
IF (uChannelCount <= 0) OR (uChannelCount > nMaxCh) THEN
    bCfgFault := TRUE;                    // 组态非法：全输出维持 FALSE（段 1 已清）
    nErrId    := 16#0001_0201;            // 故障级：组态非法
ELSE
    bCfgFault := FALSE;                   // 解除式自证：下一拍通道数合法即解除
END_IF

(* —— 段 3：上电首拍恢复策略（仅在组态合法时生效） —— *)
IF (NOT bCfgFault) AND _bFirstScan THEN
    CASE eRestorePolicy OF

    E_DL_RestorePolicy.eHold:
        ;                                  // 保持：_abState 维持 RETAIN 语义值（上层持久化承载）
    E_DL_RestorePolicy.eReset:
        FOR _k := 0 TO (nMaxCh - 1) DO
            _abState[_k] := FALSE;         // 上电全清
        END_FOR
    E_DL_RestorePolicy.ePulse:
        FOR _k := 0 TO (nMaxCh - 1) DO
            abOut[_k] := TRUE;             // 脉冲语义：置位 1 个 PLC 周期（规格强制，防误用为持续使能）
        END_FOR
        nErrId := 16#0001_0301;            // 信息级：Pulse 上电单拍脉冲
    ELSE
        nErrId := 16#0001_0201;            // 未知恢复策略按组态错兜底（安全侧全 FALSE）
        bCfgFault := TRUE;
    END_CASE
END_IF
_bFirstScan := FALSE;                     // 首拍标志自清

(* —— 段 4：三模式解算（组态合法才执行） —— *)
IF NOT bCfgFault THEN
    CASE eMode OF

    E_DL_BtnMode.eToggle:
        FOR _k := 0 TO (uChannelCount - 1) DO
            IF artBtn[_k].Q THEN
                _abState[_k] := NOT _abState[_k];   // 单按钮翻转锁存
            END_IF
            abOut[_k] := _abState[_k];              // 输出锁存态
        END_FOR

    E_DL_BtnMode.eSingleAct:
        FOR _k := 0 TO (uChannelCount - 1) DO
            abOut[_k] := abBtn[_k];                 // 点动直通：输出 = 按钮实时电平，松开即断
        END_FOR

    E_DL_BtnMode.eSelector3:
        FOR _k := 0 TO (uChannelCount - 1) DO
            IF abBtn[_k] THEN
                IF nActiveChannel = 0 THEN
                    nActiveChannel := _k + 1;       // 记录最低按下的通道号（低通道号优先）
                ELSE
                    _bSimulKey := TRUE;             // 同拍多键：置信息码（不做静默双通）
                END_IF
            END_IF
        END_FOR
        IF _bSimulKey THEN
            nErrId := 16#0001_0101;                 // 信息级：同拍多键，低通道号优先
        END_IF
        IF nActiveChannel > 0 THEN
            FOR _k := 0 TO (uChannelCount - 1) DO
                _abState[_k] := (_k = (nActiveChannel - 1));   // 互斥：仅选中通道保持
                abOut[_k] := _abState[_k];
            END_FOR
        ELSE
            FOR _k := 0 TO (uChannelCount - 1) DO
                _abState[_k] := FALSE;              // 无键按下：互斥组全清
            END_FOR
        END_IF

    ELSE
        bCfgFault := TRUE;                          // 未知模式兜底：全 FALSE 安全侧
        nErrId := 16#0001_0201;                     // 故障级：组态非法（模式越界并入组态错）
    END_CASE
END_IF

(* —— 段 5：活动通道出口（Toggle/SingleAct 取最低活动通道） —— *)
IF (eMode = E_DL_BtnMode.eToggle) OR (eMode = E_DL_BtnMode.eSingleAct) THEN
    nActiveChannel := 0;                            // 缺省无
    FOR _k := 0 TO (uChannelCount - 1) DO
        IF abOut[_k] THEN
            nActiveChannel := _k + 1;               // 最低活动通道号
            EXIT;                                    // 找到即止
        END_IF
    END_FOR
END_IF

END_FUNCTION_BLOCK

(* ---- FB_DL_TonEx.st ---- *)
(*==============================================================================
 * 组件名称 (Component)  : FB_DL_TonEx
 * 所属子库 (Sublibrary) : DL_Base
 * 当前版本 (Version)    : 1.0.0
 * 兼容性   (Platform)   : CODESYS 3.5 / TwinCAT 3 / 汇川 InoProShop / Machine Expert
 *                         仅依赖 Standard.library（TON），零厂商方言
 * 功能描述 (Function)   : 接通延时定时器防御包装。内部委托 IEC 61131-3 标准 TON
 *                         实例完成计时内核，外围提供 PT 负值钳位与跨段输入断开
 *                         语义统一（bIN 断开当拍 ET 归零、bQ 立即 FALSE）。
 * 溯源     (Origin)     : IEC 61131-3 标准语义的道莅防御性实现
 *                         （接口语义由 IEC 61131-3 定义，clean-room 重写，
 *                         参考公开标准条款）
 * 码位     (Diag Codes) : 信息级占用区间 16#0001_014F（本件独占，仅此一码）
 *                         16#0001_014F = tPT 为负值，已钳位为 T#0s（信息级，
 *                         钳位属正常防御行为，不置故障）
 * 类型裁定 (Type Note)  : 码位段 16#0001_xxxx 为全库共享 32 位段，WORD 容量不足，
 *                         故 uDiag 采用 UDINT 承载（与库内 uErrorId : UDINT 惯例一致）
 * 依赖     (Depends)    : 无 DL_ 内部依赖；Standard.library: TON
 * 红线自检 (Redline)    : R1 ✓ 零全局变量与外部变量引用 ｜ R2 ✓ 零物理 IO 地址直写
 *                         R3 ✓ 纯 IEC 61131-3 ｜ R4 ✓ PT 钳位+除零/越界无涉
 *                         R5 ✓ 全变量中英双语同行注释 ｜ R6 N/A（无顺序状态机，见下）
 *                         R7 ✓ TON 实例主体无条件周期刷新
 * 说明     (Note)       : R6 标注 N/A —— 本组件为单步延时逻辑，不存在顺序状态机，
 *                         无 CASE 可写；非法状态不可能出现（唯一状态即"计时/直通"），
 *                         故以本节说明替代 ELSE 兜底，符合"无状态机则标注 N/A"口径。
 * 防御行为声明 (Defense): ① tPT < T#0s 时钳位为 T#0s 并置信息码 16#0001_014F
 *                           （部分平台负 TIME 行为未定义，本库统一钳 0）；
 *                         ② 跨段输入断开语义统一：bIN 断开当拍 tET 归零、bQ 立即
 *                           FALSE（由内建 TON 标准语义保证，包装层不重实现）；
 *                         ③ 首扫 bIN=TRUE 允许正常计时（TON 标准语义）但不产假 bQ
 *                           （首拍 ET 从 0 起步，bQ 天然 FALSE，无需额外抑制）。
 * 修订历史 (Revision)   :
 *   2026-11-16  v1.0.0  首版入库（R14 批 1 · T0 快车道）
 *============================================================================*)
FUNCTION_BLOCK FB_DL_TonEx
VAR_INPUT
    bIN : BOOL;   // 定时输入，TRUE 起计时，FALSE 立即复位计时 / Timing input, TRUE starts timing, FALSE resets immediately
    tPT : TIME;   // 预置延时 [ms]，负值将被钳位为 T#0s / Preset delay [ms], negative values are clamped to T#0s
END_VAR
VAR_OUTPUT
    bQ    : BOOL;   // 延时到输出，bIN 保持 TRUE 达 tPT 后置位 / Delay-elapsed output, set after bIN held TRUE for tPT
    tET   : TIME;   // 已计时 [ms]，bIN 断开当拍归零 / Elapsed time [ms], zeroed on the scan bIN drops
    uDiag : UDINT;  // 诊断字，16#0001_014F=tPT 负值已钳 0，0=无诊断事件 / Diag word, 16#0001_014F=negative tPT clamped to 0, 0=no diag event
END_VAR
VAR
    fbTon    : TON;   // 内建接通延时实例，承担计时内核 / Built-in TON instance, owns the timing kernel
    tPTClamp : TIME;  // 钳位后的预置延时 [ms]，喂给内建实例 / Clamped preset delay [ms], fed to the built-in instance
    xInit    : BOOL;  // 首扫初始化标志，FALSE=尚未完成上电初始化 / First-scan init flag, FALSE = power-on init not yet done
END_VAR

(*------------------------------------------------------------------------------
 * 段 1｜首扫初始化（历史教训⑤口径）：置于逻辑最前，禁止"初值置位后同步清零"反模式
 *      First-scan init (lesson 5): placed at the very front of the logic body
 *-----------------------------------------------------------------------------*)
IF NOT xInit THEN
    xInit    := TRUE;    // 置初始化完成标志 / Mark init as done
    tPTClamp := T#0s;    // 首扫钳位值归零，避免未初始化喂入 / Zero the clamp value on first scan, no uninitialized feed
    uDiag    := 16#0000_0000;  // 首扫诊断字清零 / Clear diag word on first scan
END_IF

(*------------------------------------------------------------------------------
 * 段 2｜PT 域校验与钳位：负 TIME 在部分平台行为未定义，统一钳 0 并置信息码；
 *      写入点排序（历史教训⑩）：本件诊断字仅有"置码 / 清码"单一分支对，无
 *      复位类与置位类竞态，排序安全
 *      PT domain check and clamp: negative TIME is undefined on some platforms,
 *      unified clamp to 0 with an informational code
 *-----------------------------------------------------------------------------*)
IF tPT < T#0s THEN
    tPTClamp := T#0s;        // 负值钳位为 0 [ms] / Clamp negative to 0 [ms]
    uDiag    := 16#0001_014F;  // 信息码：PT 负值已钳 0 / Informational: negative PT clamped to 0
ELSE
    tPTClamp := tPT;         // 域内直通 / In-domain pass-through
    uDiag    := 16#0000_0000;  // 无诊断事件，清码 / No diag event, clear code
END_IF

(*------------------------------------------------------------------------------
 * 段 3｜无条件刷新区（红线 R7）：TON 实例严禁进入任何 IF / CASE 分支；
 *      bIN 断开当拍 ET 归零、bQ 立即 FALSE 的跨段统一语义由内建 TON 标准行为保证
 *      Unconditional refresh zone (red line R7): no instance call inside IF / CASE;
 *      the unified drop-out semantics (ET zeroed and bQ FALSE on the scan bIN
 *      drops) is guaranteed by the built-in TON standard behavior
 *-----------------------------------------------------------------------------*)
fbTon(IN := bIN, PT := tPTClamp);  // 每扫描周期无条件喂入输入与钳位后 PT / Feed input and clamped PT unconditionally every scan

(*------------------------------------------------------------------------------
 * 段 4｜输出直通：bQ/tET 逐拍镜像内建实例输出，包装层不重实现计时内核
 *      Output pass-through: bQ/tET mirror the built-in outputs scan by scan;
 *      the wrapper never re-implements the timing kernel
 *-----------------------------------------------------------------------------*)
bQ  := fbTon.Q;   // 延时到输出直通 / Delay-elapsed output pass-through
tET := fbTon.ET;  // 已计时 [ms] 直通 / Elapsed time [ms] pass-through
END_FUNCTION_BLOCK

(* ---- FB_DL_TpEx.st ---- *)
(*==============================================================================
 * 组件名称 (Component)  : FB_DL_TpEx
 * 所属子库 (Sublibrary) : DL_Base
 * 当前版本 (Version)    : 1.0.0
 * 兼容性   (Platform)   : CODESYS 3.5 / TwinCAT 3 / 汇川 InoProShop / Machine Expert
 *                         仅依赖 Standard.library（TP），零厂商方言
 * 功能描述 (Function)   : 脉冲定时器防御包装。内部委托 IEC 61131-3 标准 TP 实例
 *                         完成计时内核，外围提供 PT 负值钳位，并把"不可重触发"
 *                         语义在头注释显式写死。
 * 溯源     (Origin)     : IEC 61131-3 标准语义的道莅防御性实现
 *                         （接口语义由 IEC 61131-3 定义，clean-room 重写，
 *                         参考公开标准条款）
 * 码位     (Diag Codes) : 信息级占用区间 16#0001_0151（本件独占，仅此一码）
 *                         16#0001_0151 = tPT 为负值，已钳位为 T#0s（信息级，
 *                         钳位属正常防御行为，不置故障）
 * 类型裁定 (Type Note)  : 码位段 16#0001_xxxx 为全库共享 32 位段，WORD 容量不足，
 *                         故 uDiag 采用 UDINT 承载（与库内 uErrorId : UDINT 惯例一致）
 * 依赖     (Depends)    : 无 DL_ 内部依赖；Standard.library: TP
 * 红线自检 (Redline)    : R1 ✓ 零全局变量与外部变量引用 ｜ R2 ✓ 零物理 IO 地址直写
 *                         R3 ✓ 纯 IEC 61131-3 ｜ R4 ✓ PT 钳位+除零/越界无涉
 *                         R5 ✓ 全变量中英双语同行注释 ｜ R6 N/A（无顺序状态机，见下）
 *                         R7 ✓ TP 实例主体无条件周期刷新
 * 说明     (Note)       : R6 标注 N/A —— 本组件为单步脉冲逻辑，不存在顺序状态机，
 *                         无 CASE 可写；唯一状态即"脉冲中/待触发"，以本节说明
 *                         替代 ELSE 兜底，符合"无状态机则标注 N/A"口径。
 * 防御行为声明 (Defense): ① tPT < T#0s 时钳位为 T#0s 并置信息码 16#0001_0151
 *                           （部分平台负 TIME 行为未定义，本库统一钳 0，
 *                           PT=0 时脉冲退化为单扫描周期宽度）；
 *                         ② 不可重触发语义显式化（IEC TP 标准语义，多平台实现
 *                           有偏差，此处以标准实例写死）：计时进行中 bIN 再次
 *                           触发不延长、不重启当前脉冲，必须等当前脉冲结束；
 *                         ③ R24 教训落实：本件不存在任何"实例调用前的自清/
 *                           复位写入"——段 2 钳位仅写钳位值与诊断字（纯输入域
 *                           逻辑，不触内建实例状态），实例调用后到输出镜像之间
 *                           零状态写入，bQ 不可能被前置自清压成恒 FALSE。
 * 修订历史 (Revision)   :
 *   2026-11-16  v1.0.0  首版入库（R14 批 2 · T0 快车道）
 *============================================================================*)
FUNCTION_BLOCK FB_DL_TpEx
VAR_INPUT
    bIN : BOOL;   // 触发输入，上升沿启动脉冲，计时中再触发不重启 / Trigger input, rising edge starts the pulse, retrigger during timing is ignored
    tPT : TIME;   // 脉冲宽度 [ms]，负值将被钳位为 T#0s / Pulse width [ms], negative values are clamped to T#0s
END_VAR
VAR_OUTPUT
    bQ    : BOOL;   // 脉冲输出，触发后保持 tPT 宽度 / Pulse output, held TRUE for tPT after trigger
    tET   : TIME;   // 已计时 [ms]，脉冲结束后归零 / Elapsed time [ms], zeroed after the pulse finishes
    uDiag : UDINT;  // 诊断字，16#0001_0151=tPT 负值已钳 0，0=无诊断事件 / Diag word, 16#0001_0151=negative tPT clamped to 0, 0=no diag event
END_VAR
VAR
    fbTp     : TP;    // 内建脉冲定时器实例，承担计时内核 / Built-in TP instance, owns the timing kernel
    tPTClamp : TIME;  // 钳位后的脉冲宽度 [ms]，喂给内建实例 / Clamped pulse width [ms], fed to the built-in instance
    xInit    : BOOL;  // 首扫初始化标志，FALSE=尚未完成上电初始化 / First-scan init flag, FALSE = power-on init not yet done
END_VAR

(*------------------------------------------------------------------------------
 * 段 1｜首扫初始化（历史教训④口径）：置于逻辑最前，首扫不产假 bQ
 *      First-scan init (lesson 4): placed at the very front, no false bQ on first scan
 *-----------------------------------------------------------------------------*)
IF NOT xInit THEN
    xInit    := TRUE;    // 置初始化完成标志 / Mark init as done
    tPTClamp := T#0s;    // 首扫钳位值归零，避免未初始化喂入 / Zero the clamp value on first scan, no uninitialized feed
    uDiag    := 16#0000_0000;  // 首扫诊断字清零 / Clear diag word on first scan
END_IF

(*------------------------------------------------------------------------------
 * 段 2｜PT 域校验与钳位（纯输入域逻辑，不触内建实例状态——R24 教训）；
 *      写入点排序审计（历史教训⑦）：本件诊断字仅有"置码/清码"单一分支对，
 *      无复位类与置位类竞态，排序安全
 *      PT domain check and clamp (input-domain only, never touches instance
 *      state - R24 lesson); single set/clear branch pair, ordering safe
 *-----------------------------------------------------------------------------*)
IF tPT < T#0s THEN
    tPTClamp := T#0s;        // 负值钳位为 0 [ms]，PT=0 脉冲退化为单拍宽度 / Clamp negative to 0 [ms], PT=0 degenerates to one-scan pulse
    uDiag    := 16#0001_0151;  // 信息码：PT 负值已钳 0 / Informational: negative PT clamped to 0
ELSE
    tPTClamp := tPT;         // 域内直通 / In-domain pass-through
    uDiag    := 16#0000_0000;  // 无诊断事件，清码 / No diag event, clear code
END_IF

(*------------------------------------------------------------------------------
 * 段 3｜无条件刷新区（红线 R7）：TP 实例严禁进入任何 IF / CASE 分支；
 *      不可重触发语义由内建标准实例行为保证，包装层零自清/复位写入，
 *      实例调用之后无任何状态写点，bQ 恒可正常动作（R24 教训）
 *      Unconditional refresh zone (red line R7): no instance call inside IF / CASE;
 *      non-retriggerable semantics is guaranteed by the built-in standard
 *      instance; zero self-clear/reset writes after the instance call
 *-----------------------------------------------------------------------------*)
fbTp(IN := bIN, PT := tPTClamp);  // 每扫描周期无条件喂入输入与钳位后 PT / Feed input and clamped PT unconditionally every scan

(*------------------------------------------------------------------------------
 * 段 4｜输出直通：bQ/tET 逐拍镜像内建实例输出，包装层不重实现计时内核
 *      Output pass-through: bQ/tET mirror the built-in outputs scan by scan;
 *      the wrapper never re-implements the timing kernel
 *-----------------------------------------------------------------------------*)
bQ  := fbTp.Q;    // 脉冲输出直通 / Pulse output pass-through
tET := fbTp.ET;   // 已计时 [ms] 直通 / Elapsed time [ms] pass-through
END_FUNCTION_BLOCK

(* ---- FB_DL_TpRetrigger.st ---- *)
(*
  ==================================================================
  组件名 Component  : FB_DL_TpRetrigger
  分类   Category   : DL_Base
  复杂度 Complexity  : cx3
  版本   Version    : 1.0.0
  功能   Purpose    : 可重触发 TP 脉冲定时变体。触发上升沿启动脉冲窗；窗内再次
                      触发沿刷新脉冲（ET 归零重启窗宽，不叠加）；窗满自动回空闲。
                      PT 钳位非负；PT=0 时 Q 为单扫描周期脉冲且 ET=0；首扫无假触发。
  来源   Source     : iec-std-wrapper（T0）
  溯源   Origin     : IEC 61131-3 标准语义的道莅防御性实现；内部委托标准 TON /
                      R_TRIG，未复制任何厂商私有库源码。
  平台   Platform   : 纯 IEC 61131-3（Standard.library: TON / R_TRIG，无私有库）
  分工声明 Split     : 与 FB_DL_PulseStretch 分工——PulseStretch 为不可重触发的
                      脉宽拉伸（首沿后窗内再沿被忽略）；本件为可重触发 TP（窗内
                      沿刷新 ET 重启窗宽），两者语义互斥，勿混用。
  作者   Author     : 道莅代码库 · PLC 编程专家（R57）
  ------------------------------------------------------------------
  边界 Boundary     :
                      一 PT 负值按信息级钳到 T#0S 执行，不锁存（每拍重算）；
                      二 重触发只刷新 ET 重启窗，不叠加窗宽；
                      三 首扫 Q 初值 FALSE，无假触发；
                      四 PT=0 时 Q 单拍脉冲且 ET=0；
                      五 无全局变量、无外部变量声明、无物理地址寻址。
  输出契约 Output contract:
                      bQ 为脉冲电平（PT=0 时退化为单拍）；bWindow 为窗活动
                      指示；tEt 为窗内流逝时间（触发拍恒为 0）；uErrorId /
                      bError 为信息级（每拍重算非锁存），锁存语义为零。
  修订记录 Revision  :
    2026-11-21  v1.0.0  R57 首版（批 1 · 序号 1）
  ==================================================================
*)

TYPE E_DL_TprPhase :
(
    eIdle  := 0,  // 空闲：无脉冲窗 / idle, no pulse window
    ePulse := 10  // 脉冲窗：窗内触发沿可重触发刷新 / pulse window, an edge inside refreshes the retrigger
);
END_TYPE

FUNCTION_BLOCK FB_DL_TpRetrigger
VAR_INPUT
    bTrig      : BOOL;            // 触发输入，上升沿启动或重触发 [-] / trigger input, a rising edge starts or retriggers
    tPulseTime : TIME := T#1S;    // 脉冲宽度 [毫秒]，负值按信息级钳零 / pulse width [millisecond], negatives clamp to zero as informational
    bEnable    : BOOL := TRUE;    // 使能，失能即清窗 [-] / enable, disabling clears the window
    bReset     : BOOL := FALSE;   // 复位上升沿清脉冲窗 [-] / reset rising edge clears the pulse window
END_VAR
VAR_OUTPUT
    bQ       : BOOL := FALSE;  // 脉冲输出 [-] / the pulse output
    bWindow  : BOOL := FALSE;  // 重触发窗活动指示 [-] / the retrigger window active indicator
    tEt      : TIME := T#0S;   // 窗内已流逝时间 [毫秒] / elapsed time inside the window [millisecond]
    uErrorId : UDINT := 0;     // 信息级码，0 = 正常 / informational code, zero is ok
    bError   : BOOL := FALSE;  // 信息级错误标志（每拍重算，非锁存）/ informational flag, recomputed each scan, not latched
END_VAR
VAR
    rtTrig   : R_TRIG; // 触发沿检测，段 0 无条件刷新 / the trigger edge, refreshed unconditionally in segment zero
    rtReset  : R_TRIG; // 复位沿检测，段 0 无条件刷新 / the reset edge, refreshed unconditionally in segment zero
    tonPulse : TON;    // 脉冲窗定时器，段 0 无条件刷新 / the pulse window timer, refreshed unconditionally
    _ePhase  : E_DL_TprPhase := E_DL_TprPhase.eIdle; // 内部相位，CASE 唯一写入目标 / internal phase, the only CASE write target
    _bActive : BOOL := FALSE; // 窗活动保持位 [-] / the window activity holder
    _tPt     : TIME := T#0S;  // 钳位后的脉冲宽度 [毫秒] / the clamped pulse width [millisecond]
END_VAR

// 段 0｜定时器与沿检测无条件周期刷新（禁入分支）；触发拍 IN 串 NOT rtTrig.Q 实现
//        单拍低电平使 TON 重启（重触发刷新 ET 的机制本体）/ segment 0, unconditional
//        refresh; the trigger scan gates IN low for one scan so the TON restarts,
//        which is the mechanism refreshing ET on a retrigger
rtTrig(CLK := bTrig); // 触发沿 / the trigger edge
rtReset(CLK := bReset); // 复位沿 / the reset edge
tonPulse(IN := _bActive AND (NOT rtTrig.Q) AND bEnable, PT := _tPt); // 脉冲窗，IN 串窗活动闸与触发拍重启闸 / the pulse window with the activity and restart gates

// 段 1｜PT 钳位非负（信息级，每拍重算不锁存）/ segment 1, PT clamped nonnegative, informational and recomputed
IF tPulseTime < T#0S THEN // 负宽度 / a negative width
    _tPt     := T#0S; // 钳到零 / clamp to zero
    uErrorId := 16#0001_0001; // 信息级：PT 负值已钳零 / informational, a negative PT clamped to zero
    bError   := TRUE; // 置信息级标志 / raise the informational flag
ELSE // 域内 / inside the domain
    _tPt     := tPulseTime; // 直通 / passthrough
    uErrorId := 16#0000_0000; // 正常码 / the ok code
    bError   := FALSE; // 信息级标志清零 / clear the informational flag
END_IF

// 段 2｜复位沿作用域：清窗保持位与相位（两项逐项声明）/ segment 2, reset edge scope declared item by item
IF rtReset.Q THEN // 复位沿 / the reset edge
    _bActive := FALSE; // 作用域一：清窗保持位 / scope one, clear the activity holder
    _ePhase  := E_DL_TprPhase.eIdle; // 作用域二：回空闲相 / scope two, back to idle
END_IF

// 段 3｜失能门控：清窗回空闲（域外行为显式，R191）/ segment 3, the disable gate, declared explicitly
IF NOT bEnable THEN // 失能 / disabled
    _bActive := FALSE; // 清窗保持位 / clear the activity holder
    _ePhase  := E_DL_TprPhase.eIdle; // 回空闲相 / back to idle
END_IF

// 段 4｜相位机：ENUM + CASE，含 ELSE 非法相位兜底（R128）/ segment 4, the phase machine with an ELSE fallback
CASE _ePhase OF

E_DL_TprPhase.eIdle: // 空闲相：等触发沿 / the idle phase, waiting for the trigger edge
    IF bEnable AND rtTrig.Q THEN // 触发沿受理（首扫沿检测自然为假，无假触发）/ the edge is accepted, no false trigger on the first scan
        _bActive := TRUE; // 开窗 / raise the window
        _ePhase  := E_DL_TprPhase.ePulse; // 迁脉冲窗相 / migrate to the pulse phase
    END_IF

E_DL_TprPhase.ePulse: // 脉冲窗相：窗内沿已在段 0 重启 TON，这里只管窗满 / the pulse phase, the restart happened in segment zero, only the expiry is handled here
    IF tonPulse.Q THEN // 窗满到期 / the window expired
        _bActive := FALSE; // 关窗 / clear the window
        _ePhase  := E_DL_TprPhase.eIdle; // 回空闲相 / back to idle
    END_IF

ELSE // 非法相位兜底（R128）/ the illegal phase fallback
    _bActive := FALSE; // 关窗 / clear the window
    _ePhase  := E_DL_TprPhase.eIdle; // 回空闲相 / back to idle
    uErrorId := 16#0001_0005; // 信息级：非法相位 / informational, an illegal phase
    bError   := TRUE; // 置信息级标志 / raise the informational flag
END_CASE

// 段 5｜统一出口：触发拍 TON 已被单拍低电平复位，故 ET=0 且 Q 立即为真 / segment 5,
//        the unified outlet; the TON was one-scan reset on the trigger scan, so ET is zero and Q rises at once
bQ      := _bActive AND (NOT tonPulse.Q) AND bEnable; // 脉冲出口（PT=0 时恰为单拍脉冲）/ the pulse outlet, a one-scan pulse when PT is zero
bWindow := _bActive AND bEnable; // 窗活动指示 / the window indicator
tEt     := tonPulse.ET; // 已流逝时间出口 / the elapsed time outlet
END_FUNCTION_BLOCK

(* ---- FB_DL_TwoHandSafety.st ---- *)
(*==============================================================================
 * 组件名称 (Component)  : FB_DL_TwoHandSafety
 * 所属子库 (Sublibrary) : DL_Base
 * 当前版本 (Version)    : 1.0.0
 * 兼容性   (Platform)   : CODESYS 3.5 / TwinCAT 3 / 汇川 InoProShop / Machine Expert
 *                         仅依赖 Standard.library（TON / R_TRIG），零厂商方言
 * 功能描述 (Function)   : 双手安全启动按钮的同步性校验与防旁路状态机。
 *                         左/右两只手按钮必须在同步窗（默认 500 ms）内先后按下才给出安全
 *                         输出；一个循环结束后必须两只手都释放才允许下一次启动；任一侧按钮
 *                         被胶带缠住、被工件压住或人为短接时，持续按下超过卡死判定时间即
 *                         升级为"旁路嫌疑"并锁存故障。典型场景是压力机、压装机、封口机——
 *                         "一只手按着启动、另一只手伸进模具"这类致死事故的全部防线。
 *                         输出侧只给一个安全位，其余全部是诊断位，避免上位机二次组合逻辑。
 *
 * 【合规披露 / Compliance disclosure（本段不得删改）】
 *   本块是标准 PLC 上的逻辑结构实现，不是安全认证功能块。ISO 13851:2019 Type IIIC
 *   要求的安全功能必须由安全继电器或安全 PLC 的安全程序承担；标准 PLC 的普通输出存在
 *   短路失效后静默失效的风险，不得作为唯一安全措施。本块的定位是：
 *   ① 在安全 PLC 中作为经过安全论证的逻辑骨架；
 *   ② 在标准 PLC 上作为非安全的工艺互锁与诊断辅助。
 *
 * 【失真披露 / Distortion disclosure】
 *   1) 输入刻意不做防抖：防抖会引入额外延时并蚕食同步窗余量，调用方必须前置
 *      FB_DL_SignalDebounce，且防抖时间计入同步窗，属串联关系而非替代关系。
 *   2) 时间判定一律用定时器 Q，不用"当前时刻减去按下时刻"，规避各平台 TIME 减法差异。
 *   3) 卡死判定跨状态持续计时：卡死按钮通常先以同步超时（0002_0001）或释放不同步
 *      （0002_0002）的面貌出现，持续计时到卡死时限后把故障码升级为 0002_0003 并置
 *      bLeftStuck/bRightStuck，HMI 才能区分"操作不规范"与"按钮被短接"。
 *
 * 开源溯源 (Origin)     : 原创实现（参考 IEC 60204-1 与 ISO 13851:2019 Type IIIC 的功能分类
 *                         与参数域，clean-room 编写，未复制任何源码）
 * 本文件内含       : TYPE  E_DL_TwoHandState（配套枚举，归属 DL_Base）
 *                    FB    FB_DL_TwoHandSafety
 * 依赖     (Depends)    : 无 DL_ 内部依赖；Standard.library: TON / R_TRIG
 * 红线自检 (Redline)    : R1 ✓ 零全局变量表与外部变量引用 ｜ R2 ✓ 零物理 IO 地址直写
 *                         R3 ✓ 纯 IEC 61131-3（无指针、无厂商私有符号）
 *                         R4 ✓ 参数钳位 + 上电锁 + 计数饱和 + 复位前提校验
 *                         R5 ✓ 全变量中英双语同行注释 ｜ R6 ✓ 五态 ENUM + CASE + ELSE 兜底
 *                         R7 ✓ 五个实例（一沿 + 四计时）主体最前部无条件刷新（本组件核心考点）
 *
 * 【取反掩码式真值约定（边界 B10）】
 *   本块接收的是"已判定为按下"的布尔量（TRUE = 按下）。现场常闭接线的按钮由调用方在
 *   硬件抽象层取反，本块不接触任何物理电平约定。
 *
 * 修订历史 (Revision)   :
 *   2026-11-14  v1.0.0  首版入库（Phase 1 收口批次 · R3）
 *============================================================================*)

(*-----------------------------------------------------------------------------
 * 枚举: E_DL_TwoHandState（归属 DL_Base，与 FB_DL_TwoHandSafety 同文件）
 * 含义: 双手安全主状态。数值步长留空位便于后续插态而不破坏已有工程。
 *----------------------------------------------------------------------------*)
TYPE E_DL_TwoHandState :
(
    eIdle        := 0,     // 待机：双手均未按下，等待首次按下 / Idle, both released
    eWaitSecond  := 10,    // 已按下单手，等待另一手在同步窗内按下 / One pressed, waiting for the second
    eBothPressed := 20,    // 双手同步按下，安全输出有效 / Both pressed synchronously, output valid
    eWaitRelease := 30,    // 已释放一手，等待另一手在释放窗内释放 / One released, waiting for the other
    eFault       := 99     // 故障锁存，仅复位沿且双手已释放可解除 / Fault latched, reset requires both released
);
END_TYPE

(*==============================================================================
 * 功能块: FB_DL_TwoHandSafety
 * 调用约定: 每个扫描周期无条件调用一次，禁止放在 IF 分支内调用。
 * 无状态泄漏: 全部状态驻留于实例私有 VAR，零全局引用，可多工位并行实例化。
 *============================================================================*)
FUNCTION_BLOCK FB_DL_TwoHandSafety
VAR_INPUT
    bLeftPressed   : BOOL;                    // 左按钮，TRUE = 按下（调用方已完成常闭取反）/ Left pressed, TRUE = pressed
    bRightPressed  : BOOL;                    // 右按钮，TRUE = 按下（调用方已完成常闭取反）/ Right pressed, TRUE = pressed
    bEnable        : BOOL := TRUE;            // 使能，FALSE 时输出立即复位且状态回待机 / Enable, FALSE drops the output and resets to idle
    tSyncWindow    : TIME := T#500MS;         // 双手同步窗 [ms]，合法域 T#0MS~500MS / Sync window [ms], valid 0..500 ms
    tReleaseWindow : TIME := T#100MS;         // 双手释放差允许窗 [ms]，合法域 T#0MS~500MS / Release difference window [ms]
    tStuckTime     : TIME := T#5S;            // 单侧持续按下判卡死时间 [s]，下限 1 s / Single-side stuck detection time [s], min 1 s
    bReset         : BOOL;                    // 上升沿：故障复位（须双手已释放）/ Rising edge: fault reset, requires both released
END_VAR
VAR_OUTPUT
    bSafeOutput    : BOOL;                    // 安全输出，仅双手同步按下期间为 TRUE / Safe output, TRUE only while both held synchronously
    bBothPressed   : BOOL;                    // 双手同时按下（无同步含义）/ Both pressed, no synchronism implied
    bSynced        : BOOL;                    // 本次启动满足同步窗 / This actuation was synchronous
    bArmed         : BOOL;                    // 已武装：自上次全部释放后尚未启动过 / Armed, no cycle since the last full release
    bLeftStuck     : BOOL;                    // 左按钮卡死嫌疑（锁存至复位）/ Left button stuck, latched until reset
    bRightStuck    : BOOL;                    // 右按钮卡死嫌疑（锁存至复位）/ Right button stuck, latched until reset
    bError         : BOOL;                    // 故障标志（锁存）/ Fault flag, latched
    uErrorId       : UDINT;                   // 故障码，0 = 无故障 / Error code, 0 = no error
    uCycleCount    : UDINT;                   // 成功完成的双手循环数（饱和）/ Completed cycles, saturating
    uAbortCount    : UDINT;                   // 同步窗前主动放弃的累计次数（饱和）/ Aborted attempts, saturating
    eState         : E_DL_TwoHandState;       // 当前状态（供 HMI 诊断）/ Current state for HMI diagnosis
END_VAR
VAR
    fbTrigReset    : R_TRIG;                  // 复位上升沿检测实例 / Reset rising edge detector
    fbTonSync      : TON;                     // 同步窗计时（单手按下期间运行）/ Sync-window timer, runs while one hand is held
    fbTonRelease   : TON;                     // 释放窗计时（另一手仍按下期间运行）/ Release-window timer, runs while the other hand stays held
    fbTonStuckL    : TON;                     // 左侧卡死计时 / Left stuck timer
    fbTonStuckR    : TON;                     // 右侧卡死计时 / Right stuck timer
    eStateInt      : E_DL_TwoHandState;       // 主状态机内部当前态 / Internal state of the main state machine
    bSyncOkLatch   : BOOL;                    // 本次启动已通过同步判定的锁存 / Latch: this actuation passed the synchronism test
    bArmLatch      : BOOL;                    // 武装标志锁存（上电必须为 FALSE）/ Armed latch, must be FALSE at power-up
    bFirstLeft     : BOOL;                    // TRUE = 本次先按下的是左手 / TRUE = the left button was pressed first
    bLeftOnly      : BOOL;                    // 仅左手按下（卡死计时的输入条件）/ Left only, the stuck-timer input condition
    bRightOnly     : BOOL;                    // 仅右手按下（卡死计时的输入条件）/ Right only, the stuck-timer input condition
    bCountCycle    : BOOL;                    // 本拍请求累加循环计数 / Cycle counter increment requested this scan
    bCountAbort    : BOOL;                    // 本拍请求累加放弃计数 / Abort counter increment requested this scan
    bCntWarned     : BOOL;                    // 计数饱和告警已发过一次 / Saturation warning already raised once
    bSkipSm        : BOOL;                    // 本拍跳过主状态机（未使能）/ Skip the state machine this scan, not enabled
    uWarnId        : UDINT;                   // 本拍瞬时告警码（参数钳位用）/ Instantaneous warning code of this scan
    bFirstScan     : BOOL := TRUE;            // 上电首扫标志 / First-scan flag
    tSyncEff       : TIME;                    // 钳位后的同步窗 [ms] / Clamped sync window [ms]
    tReleaseEff    : TIME;                    // 钳位后的释放窗 [ms] / Clamped release window [ms]
    tStuckEff      : TIME;                    // 钳位后的卡死判定时间 [ms] / Clamped stuck detection time [ms]
END_VAR
VAR CONSTANT
    DL_TH_SYNC_MAX  : TIME := T#500MS;        // 同步窗硬上限，禁止向上放宽 / Hard sync-window limit, never widened
    DL_TH_REL_MAX   : TIME := T#500MS;        // 释放窗硬上限 / Hard release-window limit
    DL_TH_STUCK_MIN : TIME := T#1S;           // 卡死判定时间下限，防正常点动误报 / Stuck-time lower bound, avoids false trips
    DL_TH_STUCK_MAX : TIME := T#1H;           // 卡死判定时间上限，防参数笔误 / Stuck-time upper bound, guards against typos
    DL_TH_CNT_MAX   : UDINT := 16#FFFF_FFFE;  // 计数器饱和值 / Counter saturation value
END_VAR

(*------------------------------------------------------------------------------
 * 段 1｜无条件刷新区（红线 R7 / 边界 B9）
 *      Unconditional refresh zone, placed at the very top of the body
 *      五个定时器的 IN 先由"状态 + 使能 + 输入组合"推导成 BOOL，实例调用本身无条件；
 *      状态取自上一拍末尾，滞后一拍是定时器语义的正常代价，换来的是永不停更
 *      IN is derived first from state and inputs; the instance call itself never sits in an IF
 *-----------------------------------------------------------------------------*)
fbTrigReset(CLK := bReset);

bLeftOnly  := bLeftPressed AND (NOT bRightPressed);
bRightOnly := bRightPressed AND (NOT bLeftPressed);

fbTonSync(IN := bEnable AND (eStateInt = E_DL_TwoHandState.eWaitSecond), PT := tSyncEff);
fbTonRelease(IN := bEnable AND (eStateInt = E_DL_TwoHandState.eWaitRelease), PT := tReleaseEff);
fbTonStuckL(IN := bEnable AND bLeftOnly, PT := tStuckEff);
fbTonStuckR(IN := bEnable AND bRightOnly, PT := tStuckEff);

(*------------------------------------------------------------------------------
 * 段 2｜上电首扫（边界 B1 的第一道防线）
 *      First-scan init: the arming latch must be FALSE, never rely on the default value
 *      上电时双手可能已被压住或短接，若武装位默认为 TRUE，第一拍就会放行
 *      A default-TRUE arming latch would release the machine on the very first scan
 *-----------------------------------------------------------------------------*)
IF bFirstScan THEN
    bFirstScan   := FALSE;
    eStateInt    := E_DL_TwoHandState.eIdle;
    bArmLatch    := FALSE;
    bSyncOkLatch := FALSE;
    bLeftStuck   := FALSE;
    bRightStuck  := FALSE;
END_IF

(*------------------------------------------------------------------------------
 * 段 3｜时间参数钳位（边界 B3/B4/B5）
 *      Parameter clamping: widening the window means weakening safety, so clamp downwards only
 *      放宽同步窗等于放宽安全，因此越上限只向下钳位并告警；下限方向同理
 *-----------------------------------------------------------------------------*)
tSyncEff    := tSyncWindow;
tReleaseEff := tReleaseWindow;
tStuckEff   := tStuckTime;
uWarnId     := 16#0000;

IF tSyncEff > DL_TH_SYNC_MAX THEN
    tSyncEff  := DL_TH_SYNC_MAX;
    uWarnId   := 16#0001_0001;
END_IF

IF tSyncEff < T#0MS THEN
    tSyncEff  := T#0MS;
    uWarnId   := 16#0001_0001;
END_IF

IF tReleaseEff > DL_TH_REL_MAX THEN
    tReleaseEff := DL_TH_REL_MAX;
    uWarnId     := 16#0001_0001;
END_IF

IF tReleaseEff < T#0MS THEN
    tReleaseEff := T#0MS;
    uWarnId     := 16#0001_0001;
END_IF

IF tStuckEff < DL_TH_STUCK_MIN THEN
    tStuckEff := DL_TH_STUCK_MIN;
    uWarnId   := 16#0001_0001;
END_IF

IF tStuckEff > DL_TH_STUCK_MAX THEN
    tStuckEff := DL_TH_STUCK_MAX;
    uWarnId   := 16#0001_0001;
END_IF

(*------------------------------------------------------------------------------
 * 段 4｜故障码口径（红线 R15）
 *      Error-code policy: a latched code survives until the reset path clears it
 *      故障锁存期间必须保留进入故障时的码，否则 HMI 下一拍读回 0，根因丢失；
 *      非故障态下瞬时告警每拍重算，条件消失即归零
 *-----------------------------------------------------------------------------*)
IF eStateInt <> E_DL_TwoHandState.eFault THEN
    IF uWarnId <> 16#0000 THEN
        uErrorId := uWarnId;
    ELSE
        uErrorId := 16#0000_0000;
    END_IF
END_IF

(*------------------------------------------------------------------------------
 * 段 5｜未使能处理：输出撤销、状态回待机、清码但不计故障
 *      Disabled: drop the output, return to idle, clear the code without recording a fault
 *      未使能是操作员的主动动作，不是故障；重新使能后仍必须重新武装才可能放行
 *-----------------------------------------------------------------------------*)
bSkipSm := FALSE;

IF NOT bEnable THEN
    eStateInt    := E_DL_TwoHandState.eIdle;
    bArmLatch    := FALSE;
    bSyncOkLatch := FALSE;
    bLeftStuck   := FALSE;
    bRightStuck  := FALSE;
    uErrorId     := 16#0000_0000;
    bSkipSm      := TRUE;
END_IF

IF NOT bSkipSm THEN

    (*--------------------------------------------------------------------------
     * 段 6｜卡死诊断（边界 B6 的对应项）：先于主状态机判定
     *      Stuck diagnosis runs before the state machine
     *      仅单侧持续按下才计时；双手同时按下属正常操作，绝不参与卡死计时
     *      卡死按钮往往先以同步超时码出现，到时后升级为旁路嫌疑码——这是 HMI 区分
     *      "操作不规范"与"按钮被短接"的唯一依据
     *      A stuck button first shows up as a sync timeout; the upgrade to the bypass code
     *      is what lets the HMI tell sloppy operation from a taped-down button
     *-------------------------------------------------------------------------*)
    IF fbTonStuckL.Q OR fbTonStuckR.Q THEN
        bLeftStuck  := bLeftStuck OR fbTonStuckL.Q;
        bRightStuck := bRightStuck OR fbTonStuckR.Q;
        eStateInt   := E_DL_TwoHandState.eFault;
        uErrorId    := 16#0002_0003;
    END_IF

    (*--------------------------------------------------------------------------
     * 段 7｜武装（边界 B1）：只有"待机且双手全释放"才武装
     *      Arming: only idle with both hands released may arm the block
     *      这是"上电时双手已被按下 / 短接"不启动的唯一保证
     *-------------------------------------------------------------------------*)
    IF (eStateInt = E_DL_TwoHandState.eIdle) AND (NOT bLeftPressed) AND (NOT bRightPressed) THEN
        bArmLatch := TRUE;
    END_IF

    bCountCycle := FALSE;
    bCountAbort := FALSE;

    (*--------------------------------------------------------------------------
     * 段 8｜主状态机（红线 R6）：ENUM + CASE + ELSE 兜底
     *      Main state machine with the mandatory ELSE fallback
     *-------------------------------------------------------------------------*)
    CASE eStateInt OF

        E_DL_TwoHandState.eIdle:
            (* 未武装时的任何按下都被忽略，状态原地不动（边界 B1） *)
            (* Without arming, any press is ignored and the state stays put *)
            IF bArmLatch AND (bLeftPressed OR bRightPressed) THEN
                bSyncOkLatch := FALSE;
                IF bLeftPressed AND bRightPressed THEN
                    (* 边界 B2：同拍按下直接判定同步成功，但仍需武装 *)
                    (* Same-scan press counts as synchronous, arming still required *)
                    bSyncOkLatch := TRUE;
                    bArmLatch    := FALSE;
                    bCountCycle  := TRUE;
                    eStateInt    := E_DL_TwoHandState.eBothPressed;
                ELSE
                    bFirstLeft := bLeftPressed;
                    eStateInt  := E_DL_TwoHandState.eWaitSecond;
                END_IF
            END_IF

        E_DL_TwoHandState.eWaitSecond:
            (* 超时优先判定：定时器 Q 是唯一依据，不做 TIME 减法 *)
            (* Timeout first: the timer Q is the only criterion, no TIME subtraction *)
            IF fbTonSync.Q THEN
                eStateInt := E_DL_TwoHandState.eFault;
                uErrorId  := 16#0002_0001;
            ELSIF bLeftPressed AND bRightPressed THEN
                bSyncOkLatch := TRUE;
                bArmLatch    := FALSE;
                bCountCycle  := TRUE;
                eStateInt    := E_DL_TwoHandState.eBothPressed;
            ELSIF (bFirstLeft AND (NOT bLeftPressed)) OR ((NOT bFirstLeft) AND (NOT bRightPressed)) THEN
                (* 先按的手先松开：本次尝试作废，不计故障但计入放弃次数 *)
                (* The first hand released: the attempt is void, counted as an abort, not a fault *)
                (* 同时撤销武装，必须重新全释放才能再来一次，防止反复空跳 *)
                (* Arming is dropped as well, a full release is required before the next attempt *)
                bArmLatch    := FALSE;
                bSyncOkLatch := FALSE;
                bCountAbort  := TRUE;
                eStateInt    := E_DL_TwoHandState.eIdle;
            END_IF

        E_DL_TwoHandState.eBothPressed:
            (* 任一手释放立即进入释放监视，输出当拍撤销（状态即输出） *)
            (* Any release starts release monitoring; the output drops within the same scan *)
            IF NOT (bLeftPressed AND bRightPressed) THEN
                eStateInt := E_DL_TwoHandState.eWaitRelease;
            END_IF

        E_DL_TwoHandState.eWaitRelease:
            (* 两只手都释放是成功路径，优先于超时判定 *)
            (* Both released is the success path and wins over the timeout *)
            IF (NOT bLeftPressed) AND (NOT bRightPressed) THEN
                eStateInt := E_DL_TwoHandState.eIdle;
                bArmLatch := FALSE;
            ELSIF fbTonRelease.Q THEN
                eStateInt := E_DL_TwoHandState.eFault;
                uErrorId  := 16#0002_0002;
            END_IF

        E_DL_TwoHandState.eFault:
            (* 边界 B6：双手未全释放时复位无效，否则"按住一手 + 复位"即可旁路 *)
            (* Reset is ignored unless both hands are released, otherwise it is a bypass *)
            IF fbTrigReset.Q AND (NOT bLeftPressed) AND (NOT bRightPressed) THEN
                eStateInt    := E_DL_TwoHandState.eIdle;
                uErrorId     := 16#0000_0000;
                bSyncOkLatch := FALSE;
                bArmLatch    := FALSE;
                bLeftStuck   := FALSE;
                bRightStuck  := FALSE;
            END_IF

        ELSE
            (* 非法状态拦截：不做隐式恢复，直接锁存上报 *)
            (* Illegal state interception: no implicit recovery, latch and report *)
            eStateInt := E_DL_TwoHandState.eFault;
            uErrorId  := 16#0001_0005;

    END_CASE;

    (*--------------------------------------------------------------------------
     * 段 9｜计数器累加（边界 B7）：单一累加点 + 饱和不再回绕
     *      Counter accumulation: one single increment point with saturation
     *      回绕会让"运行了 43 亿次"变成"0 次"，保养周期判断随之失效
     *-------------------------------------------------------------------------*)
    IF bCountCycle THEN
        IF uCycleCount < DL_TH_CNT_MAX THEN
            uCycleCount := uCycleCount + 1;
        ELSIF NOT bCntWarned THEN
            uErrorId   := 16#0001_0007;
            bCntWarned := TRUE;
        END_IF
    END_IF

    IF bCountAbort THEN
        IF uAbortCount < DL_TH_CNT_MAX THEN
            uAbortCount := uAbortCount + 1;
        ELSIF NOT bCntWarned THEN
            uErrorId   := 16#0001_0007;
            bCntWarned := TRUE;
        END_IF
    END_IF

END_IF

(*------------------------------------------------------------------------------
 * 段 10｜输出单一出口（边界 B9 / 范式 P-05）
 *      Single output exit: the safe bit is assigned exactly once, here
 *      分支内只改状态，输出全部在末尾由状态派生，杜绝"多处置位、漏撤一处"的经典事故
 *      Branches only move the state; the safe bit derives from the state in one place
 *-----------------------------------------------------------------------------*)
bSafeOutput  := (eStateInt = E_DL_TwoHandState.eBothPressed) AND bEnable;
bBothPressed := bLeftPressed AND bRightPressed;
bSynced      := bSyncOkLatch AND bEnable;
bArmed       := bArmLatch;
bError       := (eStateInt = E_DL_TwoHandState.eFault);
eState       := eStateInt;
END_FUNCTION_BLOCK

(* ---- FB_DL_TwoStepConfirm.st ---- *)
(*
  ==================================================================
  组件名 Component  : FB_DL_TwoStepConfirm
  分类   Category   : DL_Base
  复杂度 Complexity  : 中
  版本   Version    : 1.0.2
  功能   Purpose    : 两步确认防误触发。首按（上升沿）进入预备态 bArmed，
                      限窗 tArmWindow 内二按（再次上升沿）才输出确认单脉冲
                      bConfirmed；预备窗超时自动复位并输出超时单脉冲
                      bTimeout。IEC 60204 人机交互公开语义（双手/两步确认
                      防误触发思想），与 FB_DL_HoldRepeatButton 按住重复分工。
  来源   Source     : self-std（IEC 60204 公开人机交互语义）
  溯源   Origin     : IEC 60204-1 两步控制公开条款语义，clean-room 自研实现，
                      未复制任何厂商私有库源码。
  平台   Platform   : 纯 IEC 61131-3（Standard.library: TON / R_TRIG，无私有库）
  分工声明 Split     : 与 FB_DL_HoldRepeatButton 分工——后者做按住重复触发，
                      本件做两步防误确认。
  作者   Author     : 道莅代码库 · PLC 编程专家（R59）
  ------------------------------------------------------------------
  边界 Boundary     :
                      一 确认/超时均为单拍脉冲输出，每拍先统一预清零再置位
                         （本库纪律③，防粘滞）；
                      二 预备窗 tArmWindow 超时自动复位预备态（窗口末退出迁
                         移，本库纪律④）；
                      三 busy 态（已预备）期间忽略一切新输入语义，只接受二
                         按 / 超时两条出口；
                      四 定时器与沿检测全部段 0 无条件周期刷新（R7）；
                      五 段序铁律：段 3 先消化本拍输入沿、段 4 才做超时迁移，
                         窗口到期拍与二按沿同拍时二按优先，bTimeout 不在该拍
                         发码（R275 同拍竞态口径）；
                      六 无全局变量、无外部变量声明、无物理地址寻址。
  修订记录 Revision  :
    2026-11-21  v1.0.0  R59 首版（批 1 · 序号 2）
    2026-11-21  v1.0.1  修 R275 同拍竞态：超时迁移前预消化本拍二按沿
                        （原 v1.0.0 段 3 超时先清 _bArmed，段 4 读假预备态把
                         二按当首按重新武装，二按被吞需按第三次；本次仅调整
                         段序与事件优先判据，对外引脚与语义一字不动）
    2026-11-21  v1.0.2  R61 轻项：段 4 超时判据补 AND _bArmed 双保险（R60
                        复核残留项；语义不变，仅防御性收紧）
  ==================================================================
*)

FUNCTION_BLOCK FB_DL_TwoStepConfirm
VAR_INPUT
    bBtn       : BOOL := FALSE;  // 确认按钮输入，上升沿语义 [-] / the confirm button input, rising edge semantics
    tArmWindow : TIME := T#3S;   // 二按限窗时长 [毫秒] / the second press window [millisecond]
END_VAR
VAR_OUTPUT
    bArmed     : BOOL := FALSE;  // 预备态指示（首按已受理等二按）[-] / the armed indicator, first press accepted
    bConfirmed : BOOL := FALSE;  // 两步确认成立单脉冲（单拍）[-] / the confirmed one shot pulse, single scan
    bTimeout   : BOOL := FALSE;  // 预备窗超时单脉冲（单拍）[-] / the window timeout one shot pulse, single scan
    bError     : BOOL := FALSE;  // 预留故障位（本件无浮点运算，恒常假）[-] / the reserved fault bit, constant false
END_VAR
VAR
    _bInit     : BOOL := FALSE; // 首拍初始化标志（R310，真实使用：首拍清预备态）/ the first scan flag, real use
    _bArmed    : BOOL := FALSE; // 预备态锁存位（区分于实时镜像 bArmed）/ the armed latch bit
    _bEvtTaken : BOOL := FALSE; // 同拍事件已消化标志（单拍，段 2 预清，R275）/ the same scan event consumed flag, single scan preset in segment two
    rtBtn      : R_TRIG;        // 按钮沿检测，段 0 无条件刷新 / the button edge, refreshed unconditionally
    tonArm     : TON;           // 二按限窗定时器，段 0 无条件刷新 / the arm window timer, refreshed unconditionally
END_VAR

// 段 0｜定时器与沿检测无条件周期刷新（禁入分支，R7）/ segment 0, the unconditional refresh
rtBtn(CLK := bBtn); // 按钮沿 / the button edge
tonArm(IN := _bArmed, PT := tArmWindow); // 限窗计时，预备态驱动 / the window timing, driven by the armed latch

// 段 1｜首拍初始化（R310 真实使用路径）：预备态显式清零 / segment 1, the first scan init
IF NOT _bInit THEN // 首拍一拍 / the first scan
    _bInit := TRUE; // 置首拍标志 / raise the first scan flag
    _bArmed := FALSE; // 预备态显式清零（编译缺省之上的显式安全预置）/ clear the armed latch explicitly
END_IF

// 段 2｜单拍脉冲与单拍标志每拍前置清零（本库纪律③防粘滞；仅单拍标志入此清单，R32 FB32-1）/ segment 2, the per scan preset of the one shot pulses and flags
bConfirmed := FALSE; // 确认脉冲预清零 / preset the confirmed pulse false
bTimeout := FALSE; // 超时脉冲预清零 / preset the timeout pulse false
_bEvtTaken := FALSE; // 同拍事件消化标志预清零（先清后置，R53）/ preset the same scan consumed flag false, clear before set

// 段 3｜本拍输入沿预消化（R275：合法事件先于超时迁移消化，段序在段 4 之前）/ segment 3, the same scan input edge pre-digest, the legal event ahead of the timeout migration
IF rtBtn.Q THEN // 按钮上升沿 / the button rising edge
    _bEvtTaken := TRUE; // 标记本拍已消化事件（段 4 据此不再发超时）/ mark the event consumed this scan, the segment four skips the timeout
    IF NOT _bArmed THEN // 首按：进入预备 / the first press, arm
        _bArmed := TRUE; // 置预备态（限窗同步启动）/ raise the armed latch
    ELSE // 二按：确认成立 / the second press, confirmed
        _bArmed := FALSE; // 退出预备态 / leave the armed state
        bConfirmed := TRUE; // 置确认单脉冲 / raise the confirmed pulse
    END_IF
END_IF

// 段 4｜预备窗超时迁移（窗口末退出，边界二；同拍已消化输入沿则不迁移，R275）/ segment 4, the window expiry migration, skipped when the same scan edge is already consumed
IF tonArm.Q AND (NOT _bEvtTaken) AND _bArmed THEN // 限窗到期且本拍无合法事件且仍在预备态（R61 轻项：_bArmed 双保险）/ the window expired with no legal event this scan and still armed, the double guard
    _bArmed := FALSE; // 自动退出预备态 / auto leave the armed state
    bTimeout := TRUE; // 置超时单脉冲 / raise the timeout pulse
END_IF

// 段 5｜统一出口（实时镜像与锁存位同源，R191 名实双出口）/ segment 5, the unified outlet
bArmed := _bArmed; // 预备态输出 / the armed outlet
END_FUNCTION_BLOCK

(* ---- FB_DL_UnpackWordToBits.st ---- *)
(*==============================================================================
 * 组件名称 (Component)  : FB_DL_UnpackWordToBits
 * 所属子库 (Sublibrary) : DL_Base
 * 当前版本 (Version)    : 1.0.0
 * 兼容性   (Platform)   : CODESYS 3.5 / TwinCAT 3 / 汇川 InoProShop / Machine Expert
 *                         仅依赖 Standard.library（R_TRIG），零厂商方言
 * 功能描述 (Function)   : 把通信收到的 16 位状态字 WORD 解包成 16 个独立 BOOL，
 *                         支持位取反掩码（适配常闭点），并输出"整字内容变化"的
 *                         单扫描周期事件与取反后的置位总数。
 *                         位序约定：数组索引 0 → bit0（LSB）。
 *                         R_TRIG 在主体最前部无条件刷新；上周期字在输出赋值完成之后更新。
 * 开源溯源 (Origin)     : 原创实现。变化检测采用标准异或比较 + R_TRIG 上升沿，
 *                         未使用任何厂商专有解包指令。
 * 依赖     (Depends)    : 无 DL_ 内部依赖；Standard.library: R_TRIG
 * 红线自检 (Redline)    : R1 ✓ 零全局变量表与外部变量引用 ｜ R2 ✓ 零物理 IO 地址直写
 *                         R3 ✓ 纯 IEC 61131-3 ｜ R4 ✓ 上周期值更新时序 + 下标双检 + 使能语义
 *                         R5 ✓ 全变量中英双语同行注释 ｜ R6 N/A（无顺序状态机，仅边沿锁存）
 *                         R7 ✓ R_TRIG 主体最前部无条件刷新
 * 修订历史 (Revision)   :
 *   2026-11-14  v1.0.0  首版入库（Phase 1 冷启动 · Level 0 批次）
 *============================================================================*)
FUNCTION_BLOCK FB_DL_UnpackWordToBits
VAR_INPUT
    uWord       : WORD;              // 待解包的状态字，原始值 / Source status word, raw value
    uInvertMask : WORD := 16#0000;   // 位取反掩码，对应位为 1 则输出取反 / Invert mask, a 1 bit inverts the matching output
    bEnable     : BOOL := TRUE;      // 使能标志，FALSE 时所有输出位为 FALSE / Enable flag, FALSE forces all output bits FALSE
END_VAR
VAR_OUTPUT
    abBits      : ARRAY[0..15] OF BOOL;  // 解包结果，索引 0 = bit0 / Unpacked bits, index 0 = bit0
    bChanged    : BOOL;              // 整字内容变化，单扫描周期脉冲 / Word content changed, one-scan pulse
    uBitCount   : USINT;             // 当前置位总数，值域 0..16，供冗余校验 / Popcount 0..16 for redundancy check
    uErrorId    : UDINT;             // 故障码，0 = 无故障 / Error code, 0 = no error
END_VAR
VAR
    fbTrigChange : R_TRIG;           // 整字变化检测实例 / Word change detector instance
    uXorWord     : WORD;             // 本周期与上周期的差异位（原始字比较） / XOR of current and previous raw word
    uLastWord    : WORD;             // 上周期状态字，用于差异比较 / Previous word used for difference comparison
    nIndex       : INT;              // 循环索引，值域 0..15 / Loop index, range 0..15
    uOutWord     : WORD;             // 应用取反掩码后的输出字 / Output word after applying the invert mask
    uWork        : UDINT;            // 位提取用的 UDINT 工作副本 / UDINT working copy for bit extraction
    uShift       : UDINT;            // 提升到 UDINT 的移位量 / Shift amount promoted to UDINT
    nCount       : USINT;            // 临时置位计数，值域 0..16 / Temporary popcount, range 0..16
END_VAR
VAR CONSTANT
    DL_UNPACK_BIT_COUNT : INT := 16; // 解包位数，必须与数组维度严格一致 / Unpacked bit count, must equal the array dimension
END_VAR

(*------------------------------------------------------------------------------
 * 段 1｜无条件刷新区（红线 R7 / 边界 B1）：差异比较与 R_TRIG 调用均在主体最前部
 *      Unconditional refresh zone: XOR comparison and R_TRIG call stay at the very top
 *      比较对象是"原始 uWord"，取反掩码不参与比较（边界 B3）——掩码一变若参与
 *      比较，就会被误报成现场信号跳变，把组态动作伪装成过程动作
 *      Comparison uses the raw uWord; the invert mask never participates (boundary B3)
 *-----------------------------------------------------------------------------*)
uXorWord := uWord XOR uLastWord;
fbTrigChange(CLK := (uXorWord <> 16#0000));

(*------------------------------------------------------------------------------
 * 段 2｜取反掩码应用（边界 B3）：只作用于输出位，不回头影响变化检测
 *      Invert mask applies to output bits only, never feeds back into change detection
 *-----------------------------------------------------------------------------*)
uOutWord := uWord XOR uInvertMask;
uWork    := WORD_TO_UDINT(uOutWord);
nCount   := 16#00;
uErrorId := 16#0000_0000;

IF bEnable THEN
    (*--------------------------------------------------------------------------
     * 段 3｜逐位解包 + 置位统计（边界 B4/B5）
     *      Bit-by-bit unpacking plus popcount (boundaries B4/B5)
     *      统计对象是取反后的输出位，保证 HMI 看到的位与计数同源
     *      Counting uses the post-invert bits so HMI bits and count stay consistent
     *-------------------------------------------------------------------------*)
    FOR nIndex := 0 TO (DL_UNPACK_BIT_COUNT - 1) DO
        IF (nIndex >= 0) AND (nIndex <= (DL_UNPACK_BIT_COUNT - 1)) THEN
            uShift := INT_TO_UDINT(nIndex);
            IF (SHR(uWork, uShift) AND 16#0000_0001) <> 16#0000_0000 THEN
                abBits[nIndex] := TRUE;
                nCount         := nCount + 16#01;
            ELSE
                abBits[nIndex] := FALSE;
            END_IF
        ELSE
            (* 下标越界兜底：理论上不可达（循环上界即数组上界），仍显式上报 *)
            (* Index out-of-range fallback: unreachable in theory, still reported explicitly *)
            uErrorId := 16#0001_0007;
        END_IF
    END_FOR;

    uBitCount := nCount;

    (* 变化事件：仅在使能时对外可见，禁用期间的差异由 uLastWord 继续跟踪吸收 *)
    (* Change event is visible only while enabled, differences while disabled are absorbed *)
    bChanged := fbTrigChange.Q;
ELSE
    (*--------------------------------------------------------------------------
     * 段 4｜使能失效语义（边界 B6）：输出位全 FALSE、计数清零
     *      Disabled: all output bits FALSE and the popcount cleared
     *-------------------------------------------------------------------------*)
    FOR nIndex := 0 TO (DL_UNPACK_BIT_COUNT - 1) DO
        IF (nIndex >= 0) AND (nIndex <= (DL_UNPACK_BIT_COUNT - 1)) THEN
            abBits[nIndex] := FALSE;
        END_IF
    END_FOR;

    uBitCount := 16#00;
    bChanged  := FALSE;
END_IF

(*------------------------------------------------------------------------------
 * 段 5｜上周期字更新（边界 B2，硬性顺序）：必须在输出赋值完成之后
 *      Previous word update: must happen strictly after the outputs are assigned
 *      若提前到段 1 之前或之中，异或结果恒为 0，变化事件将永久失效
 *-----------------------------------------------------------------------------*)
uLastWord := uWord;
END_FUNCTION_BLOCK

(* ---- FB_DL_ValueHoldMonitor.st ---- *)
(*
  FB_DL_ValueHoldMonitor  —  信号冻结保持监视：域外/超时保持最后有效值 + 掩码标记 / Value hold monitor with mask flags
  分类 Category : DL_Base
  版本 Version  : 1.0.0
  来源 Source   : t1-2-oscat — 域外显式化纪律零检索深化
  溯源 Origin   : clean-room 实现，未复制任何源码行
  功能 Function : 1) 输入域外或冻结超时 → 输出保持最后有效值 fHoldVal，掩码 uMask 置位
                  （bit0 = 域外，bit1 = 超时冻结），恢复输出须域内连续 nConfirm 拍；
                  2) 域判据全部使用当拍量（fIn 与组态引脚），无锁存量自指；
                  3) 掩码位序与故障码一一对应：域外→04A8、超时→04A9；
                  4) 域外/超时为保持态（故障级 03E5 锁存至 bReset），恢复且复位后清。
  边界 Boundary : ① 组态闸：fLoLim < fHiLim、nConfirm >= 1、fChgTol >= 0 必须成立，
                  违例置故障级 03E4，输出冻结为最后有效值；
                  ② 保持相 CASE 全覆盖 + ELSE 兜底落 03E6；
                  ③ 恢复计数仅在域内且非冻结拍递增，域外即清零；
                  ④ 无 GVL 依赖：纯引脚输入输出，无外部变量引用，无物理 IO 地址。
  依赖 Depends  : 仅 Standard.library（TON / R_TRIG）
  码表 Error codes（Base 段 0001，窗口 03E4~03E6 / 04A7~04A9）:
    16#0001_03E4 故障级：组态非法（量程颠倒 / nConfirm < 1 / 容差为负），锁存至 bReset
    16#0001_03E5 故障级：信号保持激活（域外或冻结超时），锁存至 bReset + 域内恢复
    16#0001_03E6 故障级：保持相位落 ELSE 兜底（非法相位 ID），锁存至 bReset
    16#0001_04A7 信息级：新值恢复确认（nConfirm 拍域内沿）
    16#0001_04A8 信息级：域外检出（伴随态，掩码 bit0）
    16#0001_04A9 信息级：冻结超时检出（伴随态，掩码 bit1）
  修订历史 Revision :
    2026-11-19  v1.0.0  R41 首版（批次 2 · 序号 1）
*)

TYPE E_DL_VhmState :
(
    eLive := 0,    // 实时透传：输出跟随输入 / Live, output follows the input
    eHold := 10,   // 保持：输出冻结最后有效值 / Hold, output frozen to last valid value
    eConf := 20    // 恢复确认：域内连续计数中 / Confirm, counting in-domain scans
);
END_TYPE

FUNCTION_BLOCK FB_DL_ValueHoldMonitor
VAR_INPUT
    fIn          : LREAL := 0.0;      // 被监视输入 [EU] / Monitored input
    fLoLim       : LREAL := -100.0;   // 有效域下限 [EU]，必须 < fHiLim / Valid span lower bound
    fHiLim       : LREAL := 100.0;    // 有效域上限 [EU]，必须 > fLoLim / Valid span upper bound
    fChgTol      : LREAL := 1.0E-6;   // 冻结判定容差 [EU]，域 >= 0 / Freeze tolerance on change
    tHoldTo      : TIME := T#5S;      // 冻结确认超时 [ms]，域 > 0 / Freeze confirm timeout
    nConfirm     : INT := 3;          // 恢复确认拍数 [拍]，域 >= 1 / Recovery confirm scans
    bReset       : BOOL := FALSE;     // 复位，上升沿清故障锁存 / Reset edge clears fault latch
END_VAR
VAR_OUTPUT
    fOut         : LREAL;             // 输出：实时值或保持值 [EU] / Output: live or held value
    bHeld        : BOOL;              // 保持中标志 [-] / Holding flag
    uMask        : WORD;              // 掩码：bit0 域外 / bit1 超时冻结 / Mask flags
    bValid       : BOOL;              // 输出有效（实时相 TRUE）/ Output usable flag
    bError       : BOOL;              // 故障锁存标志 / Fault latch flag
    nErrId       : UDINT;             // 事件码，0 = 无事件 / Event code
END_VAR
VAR
    tonHoldTo    : TON;               // 冻结确认定时器，无条件周期刷新 / Freeze confirm timer
    rtReset      : R_TRIG;            // 复位沿实例，无条件周期刷新 / Reset edge instance
    _eState      : E_DL_VhmState := E_DL_VhmState.eLive;  // 内部相位（CASE 唯一写入目标）/ Internal phase
    _fHoldVal    : LREAL := 0.0;      // 最后有效值快照 [EU] / Last valid value snapshot
    _nConfCnt    : INT;               // 恢复确认计数 [拍] / Recovery confirm counter
    _bInDom      : BOOL;              // 域内判定（当拍量）/ In-domain current-scan flag
    _bFault      : BOOL;              // 故障锁存位（锁存量）/ Latched fault bit
    _uFault      : UDINT;             // 故障码锁存（锁存量）/ Latched fault code
    _uInfo       : UDINT;             // 信息码，每拍重算 / Transient info code
    _bLivePrev   : BOOL;              // 上拍实时相镜像（恢复沿判据）/ Previous live mirror
END_VAR

(* —— 段 0：定时器与沿实例无条件周期刷新（禁置于 IF/CASE 内） —— *)
_bInDom := (fIn >= fLoLim) AND (fIn <= fHiLim);         // 域内判定（当拍量）
tonHoldTo(IN := (ABS(fIn - _fHoldVal) <= fChgTol), PT := tHoldTo);  // 冻结确认（每拍必调）
rtReset(CLK := bReset);                                 // 复位沿（每拍必调）

(* —— 段 1：单拍量预清零（锁存量 _bFault/_uFault/_fHoldVal 不入清单，禁同拍抹除） —— *)
_uInfo := 16#0000_0000;             // 信息码每拍重算
uMask := 16#0000;                   // 掩码每拍重算
bValid := FALSE;                    // 有效出口缺省 FALSE
nErrId := 16#0000_0000;             // 事件码缺省无事件

(* —— 段 2：复位沿（唯一故障解除路径，全当拍量） —— *)
IF rtReset.Q THEN                   // rtReset.Q = 当拍量
    _bFault := FALSE;               // 清故障锁存位
    _uFault := 16#0000_0000;        // 清故障锁存码
END_IF

(* —— 段 3：组态域闸（覆盖参与判据换算的全部组态引脚） —— *)
IF (fLoLim >= fHiLim) OR (nConfirm < 1) OR (fChgTol < 0.0) OR (TIME_TO_DINT(tHoldTo) <= 0) THEN
    _uFault := 16#0001_03E4;        // 故障级：组态非法
    _bFault := TRUE;
END_IF

(* —— 段 4：保持相位机（CASE 全覆盖 + ELSE 兜底） —— *)
CASE _eState OF

E_DL_VhmState.eLive:
    IF NOT _bInDom THEN
        uMask := uMask OR 16#0001;      // 掩码 bit0：域外
        _uInfo := 16#0001_04A8;         // 信息级：域外检出
        _eState := E_DL_VhmState.eHold; // 进保持相
    ELSIF tonHoldTo.Q THEN
        uMask := uMask OR 16#0002;      // 掩码 bit1：超时冻结
        _uInfo := 16#0001_04A9;         // 信息级：冻结超时
        _eState := E_DL_VhmState.eHold; // 进保持相
    ELSE
        _fHoldVal := fIn;               // 实时相刷新最后有效值快照
    END_IF

E_DL_VhmState.eHold:
    uMask := uMask OR 16#0001;          // 保持相：掩码 bit0 维持（域外/超时聚合保持）
    IF tonHoldTo.Q THEN
        uMask := uMask OR 16#0002;      // 掩码 bit1：冻结持续
    END_IF
    IF _bInDom AND (NOT tonHoldTo.Q) THEN
        _nConfCnt := 0;                 // 域内首拍：确认计数清零起步
        _eState := E_DL_VhmState.eConf; // 进恢复确认相
    END_IF

E_DL_VhmState.eConf:
    IF _bInDom AND (NOT tonHoldTo.Q) THEN
        _nConfCnt := _nConfCnt + 1;     // 域内连续计数递增
        IF _nConfCnt >= nConfirm THEN
            _uInfo := 16#0001_04A7;     // 信息级：新值恢复确认沿
            _eState := E_DL_VhmState.eLive;  // 回实时透传相
        END_IF
    ELSE
        _nConfCnt := 0;                 // 域外即清零
        _eState := E_DL_VhmState.eHold; // 回保持相
    END_IF

ELSE
    _uFault := 16#0001_03E6;        // 故障级：非法相位 ID 兜底
    _bFault := TRUE;
    _eState := E_DL_VhmState.eHold; // 强制回保持相（安全侧）

END_CASE

(* —— 段 5：保持聚合故障锁存（03E5：保持态持续或组态闸；解除 = 复位沿 + 恢复确认） —— *)
IF (_eState <> E_DL_VhmState.eLive) OR _bFault THEN
    IF NOT _bFault THEN
        _uFault := 16#0001_03E5;    // 故障级：信号保持激活（首次进入锁存）
    END_IF
    _bFault := TRUE;                // 锁存位维持（恢复相不自动清，须复位沿）
END_IF

(* —— 段 6：出口单点映射（名实同源；锁存码回放，禁同拍抹除） —— *)
IF _eState = E_DL_VhmState.eLive THEN
    fOut := fIn;                    // 实时透传
    bValid := NOT _bFault;          // 有效出口（故障期保持 FALSE）
ELSE
    fOut := _fHoldVal;              // 保持最后有效值
    bValid := FALSE;                // 保持相输出不可用
END_IF
bHeld := (_eState <> E_DL_VhmState.eLive);   // 保持中派生位
IF _bFault THEN
    nErrId := _uFault;              // 故障锁存码回放
ELSE
    nErrId := _uInfo;               // 信息码
END_IF
bError := _bFault;                  // 故障标志与锁存位同源
_bLivePrev := (_eState = E_DL_VhmState.eLive);  // 恢复沿判据快照

END_FUNCTION_BLOCK
